(* IEC 61131-3 sources: daoli-st-library/DL_Base (part 3) *)

(* ---- FC_DL_StringRemoveWhitespace.st ---- *)
(*==============================================================================
 * 组件名称 (Component)  : FC_DL_StringRemoveWhitespace
 * 所属子库 (Sublibrary) : DL_Base
 * 当前版本 (Version)    : 1.0.0
 * 兼容性   (Platform)   : CODESYS 3.5+ / TwinCAT 3 / 汇川 InoProShop / 施耐德 Machine Expert
 *                         仅依赖 IEC 61131-3 标准字符串九函数（LEN / MID / CONCAT / FIND），零厂商私有库
 * 功能描述 (Function)   : 剔除全部空白字符（空格 0x20 / 水平制表符 0x09），压缩 HMI 报文
 *                         与条码内容（上位机常带尾随空格或制表分隔，落盘前必须净化）。
 *                         逐字符扫描，命中空白则跳过，否则追加到输出缓冲。
 *                         空白识别用字符集常量 + FIND(集合, 单字符) > 0 判定：
 *                         集合常量内含一个字面量 TAB 字符（源码直接嵌入 0x09，
 *                         不经平台转义解析，跨平台语义一致）。
 * 接口     (Interface)  : 输入 sIn 原始字符串 [-]；
 *                         输出 sOut 净化结果、uiOutLen 结果字符数 [字符]、
 *                         uiRemoved 被剔除的空白字符数 [字符]、
 *                         eErrCode 错误码（E_DL_StrWsErr）；
 *                         返回值 = bValid 净化可信标志（TRUE = sOut 可信）。
 * 边界     (Boundary)   : ① 属主边界：只剔除空格与 TAB；CR/LF 不剔除（属协议帧结构，
 *                         由 CSV 转义件负责加引号，剔除会破坏报文语义）。
 *                         ② 长度守恒校验：LEN(sIn) = uiOutLen + uiRemoved，不守恒判故障级
 *                         eInternal 并回哨兵。
 *                         ③ 全空白输入 → 输出空串、uiOutLen=0、uiRemoved=LEN(sIn)、eOk（合法）。
 *                         ④ 扫描上界取实测长度（<=255），严格有界；全索引 1 基。
 *                         ⑤ 零全局耦合（无 GVL / VAR_EXTERNAL / 物理地址）。
 * 分工声明 (Scope)      : 与 `FC_DL_StringPadLeftZeros` 分工：本件只管剔除，补位归那件；
 *                         与 `FC_DL_StringIsNumeric` 分工：净化后再做数值判定。
 * 来源标签 (Source Tag) : 原创实现（无外部代码引入）
 * 码表     (Codes)      : 本件不占用全局数字码位；出口为 BOOL + STRING + 2×UINT +
 *                         本文件内定义 enum E_DL_StrWsErr（全库唯一）。
 * 红线自检 (Redline)    : R1 ✓ 零 GVL/VAR_EXTERNAL ｜ R2 ✓ 零 %I/%Q/%M ｜ R3 ✓ 纯 IEC 61131-3
 *                         R4 ✓ 长度守恒复检 + 扫描上界钳位 + 字符集归类（无字符码强转） ｜ R5 ✓ 声明逐行同行双语注释
 *                         R6 N/A（纯函数无状态机） ｜ R7 N/A（无实例调用）
 * 修订历史 (Revision)   : 2026-11-23  v1.0.0  R77 首版（批次 B2 · 序号 6）
 * 验收向量 (Acceptance) : ① sIn=' A B '(5 字符) → sOut='AB', uiOutLen=2, uiRemoved=3, eOk, TRUE；
 *                         ② sIn='ABC' → sOut='ABC', uiOutLen=3, uiRemoved=0, eOk；
 *                         ③ sIn='   ' → sOut='', uiOutLen=0, uiRemoved=3, eOk；
 *                         ④ sIn='' → sOut='', uiOutLen=0, uiRemoved=0, eOk。
 *==============================================================================*)

(*-----------------------------------------------------------------------------
 * 枚举: E_DL_StrWsErr（空白剔除错误码，归属 DL_Base，与本件同文件，全库唯一属主）
 *----------------------------------------------------------------------------*)
TYPE E_DL_StrWsErr :
(
    eOk       := 0,   // 信息级：剔除完成 / Info: removal completed
    eInternal := 9    // 故障级：长度守恒校验失败，结果不可信 / Fault: length conservation failed, result untrustworthy
);
END_TYPE

FUNCTION FC_DL_StringRemoveWhitespace : BOOL
VAR_INPUT
    sIn : STRING(255);   // 原始字符串 [-] / Raw input string
END_VAR
VAR_OUTPUT
    sOut      : STRING(255);   // 净化结果 [-] / Sanitized result
    uiOutLen  : UINT;          // 结果字符数 [字符] / Result character count [chars]
    uiRemoved : UINT;          // 被剔除的空白字符数 [字符] / Removed whitespace character count [chars]
    eErrCode  : E_DL_StrWsErr; // 错误码出口 [-] / Error code outlet
END_VAR
VAR
    _udLen   : UDINT;        // 输入字符数（钳位后） [字符] / Input length after clamping [chars]
    _udI     : UDINT;        // 扫描位置（1 基） [-] / Scan position, 1-based
    _sCur    : STRING(255);  // 当前单字符 [-] / Current single character
    _bSkip   : BOOL;         // 当前字符是否空白 [-] / Whether current character is whitespace
    _uiDrop  : UINT;         // 剔除累加器 [字符] / Removal accumulator [chars]
END_VAR
VAR CONSTANT
    (* 空白字符集合：首个字符为空格 0x20，第二个字符为字面量 TAB 0x09（直接嵌入） *)
    (* Whitespace set: first is space 0x20, second is a literal TAB 0x09 embedded directly *)
    DL_SWS_WS_SET  : STRING(255) := '	 ';   // 空白字符集（TAB + 空格） [-] / Whitespace set, TAB plus space
    DL_SWS_LEN_MAX : UINT := 255;           // 缓冲上限（STRING(255) 契约） [字符] / Buffer ceiling [chars]
    DL_SWS_START   : UDINT := 1;            // 字符串起始位置（IEC 1 基） [-] / String start position, 1-based
    DL_SWS_ONE_LEN : UDINT := 1;            // 单字符长度常量 [字符] / Single character length constant
END_VAR

(* —— 段 0：出口预置安全值 —— *)
FC_DL_StringRemoveWhitespace := FALSE;             // 返回值预置不可信 / Return preset untrustworthy
sOut      := '';                                   // 结果哨兵空串 / Result sentinel
uiOutLen  := 0;                                    // 长度哨兵 0 / Length sentinel
uiRemoved := 0;                                    // 剔除哨兵 0 / Removal sentinel
eErrCode  := E_DL_StrWsErr.eInternal;              // 预置最严码 / Preset strictest code

(* —— 段 1：长度实测与上域钳位（缓冲可表性反算） —— *)
_udLen := LEN(sIn);                                // 输入字符数 / Input length
IF _udLen > UINT_TO_UDINT(DL_SWS_LEN_MAX) THEN
    _udLen := UINT_TO_UDINT(DL_SWS_LEN_MAX);       // 超上限钳位 / Clamp to ceiling
END_IF

(* —— 段 2：空串早退（合法零结果） —— *)
IF _udLen = 0 THEN
    eErrCode := E_DL_StrWsErr.eOk;                 // 信息级成功 / Info success
    FC_DL_StringRemoveWhitespace := TRUE;
    RETURN;
END_IF

(* —— 段 3：逐字符扫描与选择性追加 —— *)
_uiDrop := 0;                                      // 剔除累加器清零 / Clear removal accumulator
_udI    := DL_SWS_START;                           // 起算位置 1 / Start at position one
sOut    := '';                                     // 输出缓冲显式清空 / Explicitly clear output buffer
WHILE _udI <= _udLen DO
    _sCur  := MID(sIn, DL_SWS_ONE_LEN, _udI);      // 取第 i 个字符（1 基） / Take i-th character, 1-based
    _bSkip := (FIND(DL_SWS_WS_SET, _sCur) > 0);    // 命中空白集合即跳过 / Skip when hit whitespace set
    IF _bSkip THEN
        _uiDrop := _uiDrop + 1;                    // 剔除累加 / Accumulate removal
    ELSE
        sOut := CONCAT(sOut, _sCur);               // 非空白追加 / Append non-whitespace character
    END_IF
    _udI := _udI + 1;                              // 位置步进 / Advance position
END_WHILE

(* —— 段 4：长度守恒复检（输入长度 = 保留 + 剔除） —— *)
uiOutLen  := UDINT_TO_UINT(LEN(sOut));             // 结果字符数 / Result length
uiRemoved := _uiDrop;                              // 剔除字符数 / Removed count
IF (UDINT_TO_UINT(_udLen) <> (uiOutLen + uiRemoved)) THEN
    sOut      := '';                               // 守恒失败回哨兵 / Conservation failed: sentinel
    uiOutLen  := 0;
    uiRemoved := 0;
    eErrCode  := E_DL_StrWsErr.eInternal;          // 故障级码 / Fault-level code
    RETURN;                                        // 返回 FALSE 保持 / Keep return FALSE
END_IF

(* —— 段 5：成功出口 —— *)
eErrCode := E_DL_StrWsErr.eOk;                     // 信息级成功 / Info success
FC_DL_StringRemoveWhitespace := TRUE;              // 净化可信 / Sanitization trustworthy

END_FUNCTION

(* ---- FC_DL_StringRepeat.st ---- *)
(*==============================================================================
 * 组件名称 (Component)  : FC_DL_StringRepeat
 * 所属子库 (Sublibrary) : DL_Base
 * 当前版本 (Version)    : 1.0.0
 * 兼容性   (Platform)   : CODESYS 3.5+ / TwinCAT 3 / 汇川 InoProShop / 施耐德 Machine Expert
 *                         仅依赖 IEC 61131-3 标准字符串九函数（LEN / CONCAT），零厂商私有库
 * 功能描述 (Function)   : 按次数重复拼接（分隔线 "-----"、占位符 "<><><>"、缩进填充）。
 *                         先算缓冲可容最大重复次数 = 255 DIV LEN(sIn)（分母已判零，
 *                         结构性无除零），再与请求次数比较：请求超限则按最大可容次数
 *                         截断并置 bTruncated / eTruncated（信息级，结果仍可信）；
 *                         请求次数为 0 或输入空串时输出空串。
 * 接口     (Interface)  : 输入 sIn 基元字符串 [-]、uiCount 请求重复次数 [次]；
 *                         输出 sOut 拼接结果、uiOutLen 结果字符数 [字符]、
 *                         uiApplied 实际生效次数 [次]、bTruncated 截断回执、
 *                         eErrCode 错误码（E_DL_StrRepErr）；
 *                         返回值 = bValid 拼接可信标志（TRUE = sOut 可信）。
 * 边界     (Boundary)   : ① 属主边界：只做整串重复拼接，不做单字符补位（补位归
 *                         FC_DL_StringPadLeftZeros）、不做截断加标记（归 TruncEllipsis）。
 *                         ② 除零防御：先判 LEN(sIn)=0 并早退，后才做 255 DIV LEN(sIn)。
 *                         ③ 缓冲保护：结果长度恒 <= 255（生效次数 = 255 DIV 基元长度）。
 *                         ④ uiCount=0 → 输出空串、uiApplied=0、eOk（合法零次）。
 *                         ⑤ 零全局耦合（无 GVL / VAR_EXTERNAL / 物理地址）。
 * 分工声明 (Scope)      : 与 `FC_DL_StringPadLeftZeros` 分工：定长补位归那件、
 *                         次数重复归本件；与 `FC_DL_StringTruncEllipsis` 无调用关系。
 * 来源标签 (Source Tag) : 原创实现（无外部代码引入）
 * 码表     (Codes)      : 本件不占用全局数字码位；出口为 BOOL + STRING + 3×UINT +
 *                         本文件内定义 enum E_DL_StrRepErr（全库唯一）。
 * 红线自检 (Redline)    : R1 ✓ 零 GVL/VAR_EXTERNAL ｜ R2 ✓ 零 %I/%Q/%M ｜ R3 ✓ 纯 IEC 61131-3
 *                         R4 ✓ 除零前置判零 + 缓冲上限反算 + 循环次数有界 ｜ R5 ✓ 声明逐行同行双语注释
 *                         R6 N/A（纯函数无状态机） ｜ R7 N/A（无实例调用）
 * 修订历史 (Revision)   : 2026-11-23  v1.0.0  R77 首版（批次 B2 · 序号 8）
 * 验收向量 (Acceptance) : ① sIn='AB', uiCount=3 → sOut='ABABAB', uiOutLen=6, uiApplied=3,
 *                         bTruncated=FALSE, eOk, TRUE；
 *                         ② sIn='AB', uiCount=0 → sOut='', uiOutLen=0, uiApplied=0, eOk, TRUE；
 *                         ③ sIn='', uiCount=5 → sOut='', uiOutLen=0, uiApplied=0, eOk, TRUE；
 *                         ④ sIn='X'（1 字符）, uiCount=300 → 生效 255 次，sOut 长度 255,
 *                         bTruncated=TRUE, eTruncated；
 *                         ⑤ sIn='AB', uiCount=200 → 255 DIV 2 = 127 → uiApplied=127,
 *                         长度 254, bTruncated=TRUE。
 *==============================================================================*)

(*-----------------------------------------------------------------------------
 * 枚举: E_DL_StrRepErr（重复拼接错误码，归属 DL_Base，与本件同文件，全库唯一属主）
 *----------------------------------------------------------------------------*)
TYPE E_DL_StrRepErr :
(
    eOk        := 0,   // 信息级：按请求次数完成 / Info: completed as requested
    eTruncated := 1    // 信息级：超缓冲上限已按最大可容次数截断 / Info: truncated to max fitting repeat count
);
END_TYPE

FUNCTION FC_DL_StringRepeat : BOOL
VAR_INPUT
    sIn     : STRING(255);   // 基元字符串 [-] / Unit string to repeat
    uiCount : UINT;          // 请求重复次数 [次] / Requested repeat count [times]
END_VAR
VAR_OUTPUT
    sOut       : STRING(255); // 拼接结果 [-] / Concatenated result
    uiOutLen   : UINT;        // 结果字符数 [字符] / Result character count [chars]
    uiApplied  : UINT;        // 实际生效次数 [次] / Applied repeat count [times]
    bTruncated : BOOL;        // 截断回执（信息级） [-] / Truncation receipt, info level
    eErrCode   : E_DL_StrRepErr; // 错误码出口 [-] / Error code outlet
END_VAR
VAR
    _udUnitLen : UDINT;       // 基元字符数 [字符] / Unit string length [chars]
    _udMaxRep  : UDINT;       // 缓冲可容最大重复次数 [次] / Max fitting repeat count [times]
    _uiEff     : UINT;        // 生效重复次数 [次] / Effective repeat count [times]
    _uiLoop    : UINT;        // 循环计数器 [-] / Loop counter
END_VAR
VAR CONSTANT
    DL_SRE_LEN_MAX : UINT := 255;    // 缓冲上限（STRING(255) 契约） [字符] / Buffer ceiling [chars]
    DL_SRE_ONE_LEN : UDINT := 1;     // 单字符长度常量 [字符] / Single character length constant
END_VAR

(* —— 段 0：出口预置安全值 —— *)
FC_DL_StringRepeat := FALSE;                       // 返回值预置无效 / Return preset invalid
sOut       := '';                                  // 结果哨兵空串 / Result sentinel
uiOutLen   := 0;                                   // 长度哨兵 0 / Length sentinel
uiApplied  := 0;                                   // 生效次数哨兵 0 / Applied count sentinel
bTruncated := FALSE;                               // 截断回执预置无 / Truncation receipt preset false
eErrCode   := E_DL_StrRepErr.eTruncated;           // 预置最严码（本件仅信息级码） / Preset strictest code

(* —— 段 1：基元长度实测（除零防御前置：先判零后做除法） —— *)
_udUnitLen := LEN(sIn);                            // 基元字符数 / Unit length
IF _udUnitLen = 0 THEN
    eErrCode := E_DL_StrRepErr.eOk;                // 空基元合法（零结果） / Empty unit is legal, zero result
    FC_DL_StringRepeat := TRUE;                    // 结果可信 / Result trustworthy
    RETURN;                                        // 早退，彻底规避 255 DIV 0 / Early exit, avoids division by zero entirely
END_IF

(* —— 段 2：请求次数为零早退（合法零结果） —— *)
IF uiCount = 0 THEN
    eErrCode := E_DL_StrRepErr.eOk;                // 零次合法 / Zero repeats legal
    FC_DL_StringRepeat := TRUE;
    RETURN;
END_IF

(* —— 段 3：缓冲可容最大重复次数反算（分母已确非零） —— *)
_udMaxRep := UINT_TO_UDINT(DL_SRE_LEN_MAX) / _udUnitLen;  // 255 DIV 基元长度 / Integer division by unit length
IF _udMaxRep < DL_SRE_ONE_LEN THEN
    _udMaxRep := DL_SRE_ONE_LEN;                   // 基元本身已占满缓冲：至少一次 / Unit already fills buffer: at least once
END_IF

(* —— 段 4：请求次数与可容次数比较（超限则截断并回执） —— *)
IF UINT_TO_UDINT(uiCount) > _udMaxRep THEN
    _uiEff     := UDINT_TO_UINT(_udMaxRep);         // 收敛到最大可容次数 / Converge to max fitting count
    bTruncated := TRUE;                            // 截断回执 / Truncation receipt
    eErrCode   := E_DL_StrRepErr.eTruncated;       // 信息级截断码 / Info truncation code
ELSE
    _uiEff     := uiCount;                         // 按请求次数生效 / Apply requested count
    bTruncated := FALSE;
    eErrCode   := E_DL_StrRepErr.eOk;              // 信息级成功 / Info success
END_IF

(* —— 段 5：循环拼接（次数已收敛，循环严格有界） —— *)
sOut := '';                                        // 输出缓冲显式清空 / Explicitly clear output buffer
IF _uiEff > 0 THEN
    FOR _uiLoop := 1 TO _uiEff DO
        sOut := CONCAT(sOut, sIn);                 // 每次追加一个基元 / Append one unit per iteration
    END_FOR;
END_IF

(* —— 段 6：结果复检（长度 = 基元长度 × 生效次数，且不得超缓冲） —— *)
uiOutLen  := UDINT_TO_UINT(LEN(sOut));             // 实测结果长度 / Measured result length
uiApplied := _uiEff;                               // 导出生效次数 / Export applied count
IF uiOutLen > DL_SRE_LEN_MAX THEN
    sOut      := '';                               // 超缓冲回哨兵 / Over buffer: sentinel
    uiOutLen  := 0;
    uiApplied := 0;
    eErrCode  := E_DL_StrRepErr.eTruncated;        // 保持信息级码（本件无故障级码位） / Keep info-level code
    RETURN;
END_IF

FC_DL_StringRepeat := TRUE;                        // 拼接有效 / Concatenation valid

END_FUNCTION

(* ---- FC_DL_StringReverse.st ---- *)
(*==============================================================================
 * 组件名称 (Component)  : FC_DL_StringReverse
 * 所属子库 (Sublibrary) : DL_Base
 * 当前版本 (Version)    : 1.0.0
 * 兼容性   (Platform)   : CODESYS 3.5+ / TwinCAT 3 / 汇川 InoProShop / 施耐德 Machine Expert
 *                         仅依赖 IEC 61131-3 标准字符串九函数（LEN / MID / CONCAT），零厂商私有库
 * 功能描述 (Function)   : 字符串反转（回文校验 / 字节序调试 / 低位在前的编码还原）。
 *                         自尾向头逐字符取 MID(sIn,1,i) 并 CONCAT 拼接；用 WHILE
 *                         递减计数，UDINT 计数到 0 自然终止，结构上无下溢路径。
 *                         输出长度恒等于输入长度（不做任何增删）。
 * 接口     (Interface)  : 输入 sIn 原始字符串 [-]；
 *                         输出 sOut 反转结果、uiOutLen 结果字符数 [字符]、
 *                         eErrCode 错误码（E_DL_StrRevErr）；
 *                         返回值 = bValid 反转可信标志（TRUE = sOut 可信）。
 * 边界     (Boundary)   : ① 属主边界：只做整串反转，不做大小写折叠、不做子串反转。
 *                         ② 长度 > 255 时按缓冲上限 255 截断尾部（保证输出可表），
 *                         回执 eClampLen（信息级），bTruncated 置位。
 *                         ③ 空串合法，输出空串、uiOutLen=0、eOk。
 *                         ④ 计数递减用 `IF _udI > 0` 前置判定，杜绝 UDINT 0-1 下溢。
 *                         ⑤ 零全局耦合（无 GVL / VAR_EXTERNAL / 物理地址）。
 * 分工声明 (Scope)      : 与 `FC_DL_StringCompareNatural` 分工：反转只做位序重排，
 *                         不做序比较；回文判定由调用方对 sIn 与 sOut 比较完成。
 * 来源标签 (Source Tag) : 原创实现（无外部代码引入）
 * 码表     (Codes)      : 本件不占用全局数字码位；出口为 BOOL + STRING + UINT +
 *                         本文件内定义 enum E_DL_StrRevErr（全库唯一）。
 * 红线自检 (Redline)    : R1 ✓ 零 GVL/VAR_EXTERNAL ｜ R2 ✓ 零 %I/%Q/%M ｜ R3 ✓ 纯 IEC 61131-3
 *                         R4 ✓ 递减计数下溢防护 + 长度钳位 ｜ R5 ✓ 声明逐行同行双语注释
 *                         R6 N/A（纯函数无状态机） ｜ R7 N/A（无实例调用）
 * 修订历史 (Revision)   : 2026-11-23  v1.0.0  R77 首版（批次 B2 · 序号 4）
 * 验收向量 (Acceptance) : ① sIn='ABC' → sOut='CBA', uiOutLen=3, eOk, TRUE；
 *                         ② sIn='ABBA' → sOut='ABBA'（回文自反）, uiOutLen=4；
 *                         ③ sIn='' → sOut='', uiOutLen=0, eOk, TRUE；
 *                         ④ sIn='12345' → sOut='54321'。
 *==============================================================================*)

(*-----------------------------------------------------------------------------
 * 枚举: E_DL_StrRevErr（字符串反转错误码，归属 DL_Base，与本件同文件，全库唯一属主）
 *----------------------------------------------------------------------------*)
TYPE E_DL_StrRevErr :
(
    eOk       := 0,   // 信息级：反转完成 / Info: reversal completed
    eClampLen := 1    // 信息级：长度超缓冲上限已截断 / Info: length clamped to buffer ceiling
);
END_TYPE

FUNCTION FC_DL_StringReverse : BOOL
VAR_INPUT
    sIn : STRING(255);   // 原始字符串 [-] / Raw input string
END_VAR
VAR_OUTPUT
    sOut      : STRING(255);   // 反转结果 [-] / Reversed result
    uiOutLen  : UINT;          // 结果字符数 [字符] / Result character count [chars]
    bTruncated: BOOL;          // 截断回执（信息级） [-] / Truncation receipt, info level
    eErrCode  : E_DL_StrRevErr; // 错误码出口 [-] / Error code outlet
END_VAR
VAR
    _udLen : UDINT;       // 生效字符数（钳位后） [字符] / Effective character count after clamping [chars]
    _udI   : UDINT;       // 逆序扫描位置（1 基） [-] / Reverse scan position, 1-based
END_VAR
VAR CONSTANT
    DL_SRV_LEN_MAX : UINT := 255;    // 缓冲上限（STRING(255) 契约） [字符] / Buffer ceiling [chars]
    DL_SRV_ONE_LEN : UDINT := 1;     // 单字符长度常量 [字符] / Single character length constant [chars]
END_VAR

(* —— 段 0：出口预置安全值 —— *)
FC_DL_StringReverse := FALSE;                      // 返回值预置无效 / Return preset invalid
sOut       := '';                                  // 结果哨兵空串 / Result sentinel
uiOutLen   := 0;                                   // 长度哨兵 0 / Length sentinel
bTruncated := FALSE;                               // 截断回执预置无 / Truncation receipt preset false
eErrCode   := E_DL_StrRevErr.eClampLen;            // 预置最严码（本件仅信息级码） / Preset strictest code

(* —— 段 1：长度实测与上域钳位（缓冲可表性反算） —— *)
_udLen := LEN(sIn);                                // 输入字符数 / Input length
IF _udLen > UINT_TO_UDINT(DL_SRV_LEN_MAX) THEN
    _udLen     := UINT_TO_UDINT(DL_SRV_LEN_MAX);   // 超上限截断尾部 / Truncate tail beyond ceiling
    bTruncated := TRUE;                            // 截断回执 / Truncation receipt
    eErrCode   := E_DL_StrRevErr.eClampLen;        // 信息级钳位码 / Info clamp code
ELSE
    eErrCode   := E_DL_StrRevErr.eOk;              // 信息级成功 / Info success
END_IF

(* —— 段 2：空串早退（合法零结果） —— *)
IF _udLen = 0 THEN
    FC_DL_StringReverse := TRUE;                   // 空串反转合法 / Empty reversal legal
    RETURN;
END_IF

(* —— 段 3：逆序拼接（前置 >0 判定，杜绝 UDINT 下溢） —— *)
sOut := MID(sIn, DL_SRV_ONE_LEN, _udLen);          // 以末字符起头 / Start with last character
_udI := _udLen - 1;                                // 自倒数第二位起（>=1 由段 2 保证 len>=1） / Start from second last
WHILE _udI > 0 DO
    sOut := CONCAT(sOut, MID(sIn, DL_SRV_ONE_LEN, _udI));  // 逐个前置字符追加 / Append next character from tail
    _udI := _udI - 1;                              // 位置递减，条件 >0 保证不下溢 / Decrement, guarded by >0
END_WHILE

(* —— 段 4：结果复检（长度守恒） —— *)
uiOutLen := UDINT_TO_UINT(LEN(sOut));              // 实测结果长度 / Measured result length
IF uiOutLen <> UDINT_TO_UINT(_udLen) THEN
    sOut     := '';                                // 长度不守恒回哨兵 / Length not conserved: sentinel
    uiOutLen := 0;
    eErrCode := E_DL_StrRevErr.eClampLen;          // 保持信息级码（本件无故障级码位） / Keep info-level code
END_IF

FC_DL_StringReverse := TRUE;                       // 反转有效（含截断情形） / Reversal valid, truncation included

END_FUNCTION

(* ---- FC_DL_StringSplitPair.st ---- *)
(*==============================================================================
 * 组件名称 (Component)  : FC_DL_StringSplitPair
 * 所属子库 (Sublibrary) : DL_Base
 * 当前版本 (Version)    : 1.0.0
 * 兼容性   (Platform)   : CODESYS 3.5+ / TwinCAT 3 / 汇川 InoProShop / 施耐德 Machine Expert
 *                         仅依赖 IEC 61131-3 标准字符串九函数（LEN / MID / FIND），零厂商私有库
 * 功能描述 (Function)   : key=value 单对拆分（HMI 参数设置报文 "Speed=1500" 解析）。
 *                         以首个分隔符位置为界：左侧为键、右侧为值（值可含分隔符，
 *                         故只按首个分隔符切分）。缺分隔符、空键均置无效回执（返回 FALSE），
 *                         空值合法（代表「置空」语义，回执 bHasValue=FALSE 但不判故障）。
 *                         分隔符为可配字符串（默认 '='），支持 ':=' / '->' 等双字符分隔。
 * 接口     (Interface)  : 输入 sIn 待拆分字符串 [-]、sSep 分隔符（空串回落 '='）[-]；
 *                         输出 sKey 键、sValue 值、uiKeyLen 键长 [字符]、uiValueLen 值长 [字符]、
 *                         bHasValue 是否存在值段、eErrCode 错误码（E_DL_StrSplitErr）；
 *                         返回值 = bValid 拆分有效标志（TRUE = sKey/sValue 可信）。
 * 边界     (Boundary)   : ① 属主边界：只拆单对，不遍历多对、不去引号、不做类型转换。
 *                         ② 缺分隔符 → 故障级 eNoSeparator，sKey=sIn 原样、sValue=''、返回 FALSE。
 *                         ③ 分隔符在首位（空键）→ 故障级 eEmptyKey，sKey=''、sValue=右段。
 *                         ④ 分隔符在末位（空值）→ 信息级 eEmptyValue，bHasValue=FALSE、返回 TRUE。
 *                         ⑤ MID 起算位置 = 分隔符位置 + 1，且仅当剩余长度 >= 1 时才取，
 *                         结构上无 0 长度 / 0 位置取值路径。
 *                         ⑥ 零全局耦合（无 GVL / VAR_EXTERNAL / 物理地址）。
 * 分工声明 (Scope)      : 与 `FC_DL_StringCountChar` 分工：计数归那件、拆分归本件；
 *                         与 `FC_DL_StringCsvFieldEscape` 分工：CSV 转义归那件。
 * 来源标签 (Source Tag) : 原创实现（无外部代码引入）
 * 码表     (Codes)      : 本件不占用全局数字码位；出口为 BOOL + 2×STRING + 2×UINT +
 *                         本文件内定义 enum E_DL_StrSplitErr（全库唯一）。
 * 红线自检 (Redline)    : R1 ✓ 零 GVL/VAR_EXTERNAL ｜ R2 ✓ 零 %I/%Q/%M ｜ R3 ✓ 纯 IEC 61131-3
 *                         R4 ✓ 分隔符缺失/空键域闸 + 取值位置下限保护 ｜ R5 ✓ 声明逐行同行双语注释
 *                         R6 N/A（纯函数无状态机） ｜ R7 N/A（无实例调用）
 * 修订历史 (Revision)   : 2026-11-23  v1.0.0  R77 首版（批次 B2 · 序号 7）
 * 验收向量 (Acceptance) : ① sIn='Speed=1500', sSep='=' → sKey='Speed', sValue='1500',
 *                         uiKeyLen=5, uiValueLen=4, bHasValue=TRUE, eOk, TRUE；
 *                         ② sIn='Speed1450', sSep='=' → bFound 无效：返回 FALSE, eNoSeparator, sValue=''；
 *                         ③ sIn='=1500' → 返回 FALSE, eEmptyKey, sKey='';
 *                         ④ sIn='Speed=' → sKey='Speed', sValue='', bHasValue=FALSE,
 *                         返回 TRUE, eEmptyValue；
 *                         ⑤ sIn='A=B=C' → sKey='A', sValue='B=C'（只按首个分隔符切分）；
 *                         ⑥ sIn='', sSep='=' → 返回 FALSE, eNoSeparator。
 *==============================================================================*)

(*-----------------------------------------------------------------------------
 * 枚举: E_DL_StrSplitErr（key=value 拆分错误码，归属 DL_Base，与本件同文件，全库唯一属主）
 * 分级: eEmptyValue 为信息级（返回 TRUE）；eNoSeparator / eEmptyKey 为故障级（返回 FALSE）。
 *----------------------------------------------------------------------------*)
TYPE E_DL_StrSplitErr :
(
    eOk          := 0,   // 信息级：键值均非空，拆分完成 / Info: both key and value non-empty
    eEmptyValue  := 1,   // 信息级：值段为空（置空语义） / Info: empty value section
    eNoSeparator := 2,   // 故障级：未找到分隔符 / Fault: separator not found
    eEmptyKey    := 3    // 故障级：分隔符在首位，键为空 / Fault: separator at head, empty key
);
END_TYPE

FUNCTION FC_DL_StringSplitPair : BOOL
VAR_INPUT
    sIn  : STRING(255);   // 待拆分字符串 [-] / String to split
    sSep : STRING(255);   // 分隔符（空串回落 '='） [-] / Separator, empty falls back to '='
END_VAR
VAR_OUTPUT
    sKey       : STRING(255); // 键段 [-] / Key section
    sValue     : STRING(255); // 值段 [-] / Value section
    uiKeyLen   : UINT;        // 键字符数 [字符] / Key character count [chars]
    uiValueLen : UINT;        // 值字符数 [字符] / Value character count [chars]
    bHasValue  : BOOL;        // 是否存在值段 [-] / Whether value section exists
    eErrCode   : E_DL_StrSplitErr; // 错误码出口 [-] / Error code outlet
END_VAR
VAR
    _sSepUse  : STRING(255);  // 生效分隔符 [-] / Effective separator
    _udLen    : UDINT;        // 输入字符数（钳位后） [字符] / Input length after clamping [chars]
    _udPos    : UDINT;        // 分隔符位置（1 基，0 = 未找到） [-] / Separator position, 0 means not found
    _udRemain : UDINT;        // 分隔符右侧剩余字符数 [字符] / Remaining characters after separator [chars]
    _udStart  : UDINT;        // 值段起算位置（1 基） [-] / Value section start position, 1-based
END_VAR
VAR CONSTANT
    DL_SSP_SEP_DFLT : STRING(255) := '=';   // 默认分隔符 [-] / Default separator
    DL_SSP_LEN_MAX  : UINT := 255;          // 缓冲上限（STRING(255) 契约） [字符] / Buffer ceiling [chars]
    DL_SSP_START    : UDINT := 1;           // 字符串起始位置（IEC 1 基） [-] / String start position, 1-based
END_VAR

(* —— 段 0：出口预置安全值 —— *)
FC_DL_StringSplitPair := FALSE;                    // 返回值预置无效 / Return preset invalid
sKey       := '';                                  // 键哨兵空串 / Key sentinel
sValue     := '';                                  // 值哨兵空串 / Value sentinel
uiKeyLen   := 0;                                   // 键长哨兵 0 / Key length sentinel
uiValueLen := 0;                                   // 值长哨兵 0 / Value length sentinel
bHasValue  := FALSE;                               // 值段存在性预置无 / Value presence preset false
eErrCode   := E_DL_StrSplitErr.eNoSeparator;       // 预置最严码 / Preset strictest code

(* —— 段 1：分隔符归一（空串回落默认 '='） —— *)
IF LEN(sSep) = 0 THEN
    _sSepUse := DL_SSP_SEP_DFLT;                   // 回落默认分隔符 / Fall back to default separator
ELSE
    _sSepUse := sSep;                              // 使用调用方给定分隔符 / Use caller-supplied separator
END_IF

(* —— 段 2：输入长度实测与上域钳位 —— *)
_udLen := LEN(sIn);                                // 输入字符数 / Input length
IF _udLen > UINT_TO_UDINT(DL_SSP_LEN_MAX) THEN
    _udLen := UINT_TO_UDINT(DL_SSP_LEN_MAX);       // 超上限钳位 / Clamp to ceiling
END_IF

(* —— 段 3：定位首个分隔符（FIND 返回 0 表示未找到） —— *)
_udPos := FIND(sIn, _sSepUse);                     // 首个分隔符位置（1 基） / First separator position, 1-based

(* —— 段 4：缺分隔符早退（故障级：整体原样回键，值置空） —— *)
IF _udPos = 0 THEN
    sKey     := sIn;                               // 原样回键便于调用方诊断 / Echo input to key for diagnosis
    uiKeyLen := UDINT_TO_UINT(LEN(sKey));          // 键长实测 / Measured key length
    sValue   := '';                                // 值置空 / Value cleared
    eErrCode := E_DL_StrSplitErr.eNoSeparator;     // 故障级码 / Fault-level code
    RETURN;                                        // 返回 FALSE 保持 / Keep return FALSE
END_IF

(* —— 段 5：空键闸（分隔符在首位） —— *)
IF _udPos = DL_SSP_START THEN
    sKey     := '';                                // 键为空 / Empty key
    _udRemain := _udLen - _udPos;                  // 右侧剩余长度 / Remaining length on the right
    IF _udRemain >= DL_SSP_START THEN
        sValue     := MID(sIn, _udRemain, _udPos + DL_SSP_START);  // 取分隔符之后全部字符 / Take all after separator
        uiValueLen := UDINT_TO_UINT(_udRemain);
        bHasValue  := TRUE;
    END_IF
    eErrCode := E_DL_StrSplitErr.eEmptyKey;        // 故障级码 / Fault-level code
    RETURN;                                        // 返回 FALSE 保持 / Keep return FALSE
END_IF

(* —— 段 6：键段提取（位置 1 起，长度 = 分隔符位置 - 1 >= 1） —— *)
sKey     := MID(sIn, _udPos - DL_SSP_START, DL_SSP_START);   // 分隔符左侧 / Left of separator
uiKeyLen := UDINT_TO_UINT(LEN(sKey));              // 键长实测 / Measured key length

(* —— 段 7：值段提取（起算位置 = 分隔符位置 + 1，仅剩余 >= 1 时取） —— *)
_udRemain := _udLen - _udPos;                      // 右侧剩余长度 / Remaining length on the right
IF _udRemain >= DL_SSP_START THEN
    _udStart   := _udPos + DL_SSP_START;           // 值段起算位置 / Value start position
    sValue     := MID(sIn, _udRemain, _udStart);   // 取右侧全部字符 / Take all characters on the right
    uiValueLen := UDINT_TO_UINT(LEN(sValue));      // 值长实测 / Measured value length
    bHasValue  := TRUE;                            // 存在值段 / Value section exists
    eErrCode   := E_DL_StrSplitErr.eOk;            // 信息级成功 / Info success
ELSE
    sValue     := '';                              // 分隔符在末位：值段为空 / Separator at tail: empty value
    uiValueLen := 0;
    bHasValue  := FALSE;
    eErrCode   := E_DL_StrSplitErr.eEmptyValue;    // 信息级：置空语义 / Info: clear semantics
END_IF

(* —— 段 8：键长复检（键不得为空，否则判内部不一致） —— *)
IF uiKeyLen = 0 THEN
    sKey     := '';                                // 回哨兵 / Back to sentinel
    sValue   := '';
    eErrCode := E_DL_StrSplitErr.eEmptyKey;        // 故障级码 / Fault-level code
    RETURN;
END_IF

FC_DL_StringSplitPair := TRUE;                     // 拆分有效 / Split valid

END_FUNCTION

(* ---- FC_DL_StringTruncEllipsis.st ---- *)
(*==============================================================================
 * 组件名称 (Component)  : FC_DL_StringTruncEllipsis
 * 所属子库 (Sublibrary) : DL_Base
 * 当前版本 (Version)    : 1.0.0
 * 兼容性   (Platform)   : CODESYS 3.5+ / TwinCAT 3 / 汇川 InoProShop / 施耐德 Machine Expert
 *                         仅依赖 IEC 61131-3 标准字符串九函数（LEN / MID / CONCAT），零厂商私有库
 * 功能描述 (Function)   : 超长截断并补省略标记（HMI 单行显示 / 报警摘要压缩）。
 *                         sIn 长度不超过 uiMaxLen 时原样返回；超长时保留前
 *                         (uiMaxLen - LEN(sMark)) 个字符并追加省略标记，最终长度
 *                         恒等于 uiMaxLen（标记有余量时）；标记本身已占满目标长度时
 *                         退化为纯截断（无标记空间）并回执 eTruncNoMark。
 *                         返回实际写入字符数 uiOutLen，供调用方做定宽对齐。
 * 接口     (Interface)  : 输入 sIn 原始字符串 [-]、uiMaxLen 目标最大长度（含标记）[字符]、
 *                         sMark 省略标记（空串则纯截断）[-]；
 *                         输出 sOut 结果字符串、uiOutLen 实际字符数 [字符]、
 *                         bTruncated 截断回执、eErrCode 错误码（E_DL_StrTruncErr）；
 *                         返回值 = bValid 输出可信标志（TRUE = sOut 可信）。
 * 边界     (Boundary)   : ① 属主边界：只做截断 + 单标记追加，不做补位、不剔除空白。
 *                         ② uiMaxLen 合法域 1..255；> 255 钳位至 255 并置 eClampLen；
 *                         < 1 判故障级 eInvalidParam（无法产出有效结果）。
 *                         ③ 标记长度 >= uiMaxLen 时无标记余量，退化为 MID(sIn,uiMaxLen,1)
 *                         纯截断，回执 eTruncNoMark（信息级）。
 *                         ④ 全索引 1 基，截断起算位置恒 >= 1（keep >= 1 由分支保证）。
 *                         ⑤ 零全局耦合（无 GVL / VAR_EXTERNAL / 物理地址）。
 * 分工声明 (Scope)      : 与 `FC_DL_StringPadLeftZeros` 分工：补位归那件、截断归本件，
 *                         两件互不调用；与 `FC_DL_StringRepeat` 无交集。
 * 来源标签 (Source Tag) : 原创实现（无外部代码引入）
 * 码表     (Codes)      : 本件不占用全局数字码位；出口为 BOOL + STRING + UINT +
 *                         本文件内定义 enum E_DL_StrTruncErr（全库唯一）。
 * 红线自检 (Redline)    : R1 ✓ 零 GVL/VAR_EXTERNAL ｜ R2 ✓ 零 %I/%Q/%M ｜ R3 ✓ 纯 IEC 61131-3
 *                         R4 ✓ 长度域闸 + 双侧钳位 + 起算位置下限保证 ｜ R5 ✓ 声明逐行同行双语注释
 *                         R6 N/A（纯函数无状态机） ｜ R7 N/A（无实例调用）
 * 修订历史 (Revision)   : 2026-11-23  v1.0.0  R77 首版（批次 B2 · 序号 2）
 * 验收向量 (Acceptance) : ① sIn='ABCDEFGH'（8 字符）, uiMaxLen=6, sMark='...' →
 *                         keep=3 → sOut='ABC...'（6 字符）, uiOutLen=6, bTruncated=TRUE, eOk；
 *                         ② sIn='ABC', uiMaxLen=6 → sOut='ABC'（原样）, uiOutLen=3,
 *                         bTruncated=FALSE, eOk；
 *                         ③ sIn='ABCDEFGH', uiMaxLen=3, sMark='...' → 标记占满 →
 *                         sOut='ABC', uiOutLen=3, bTruncated=TRUE, eTruncNoMark；
 *                         ④ uiMaxLen=0 → 返回 FALSE, sOut='', eInvalidParam。
 *==============================================================================*)

(*-----------------------------------------------------------------------------
 * 枚举: E_DL_StrTruncErr（截断错误码，归属 DL_Base，与本件同文件，全库唯一属主）
 *----------------------------------------------------------------------------*)
TYPE E_DL_StrTruncErr :
(
    eOk           := 0,   // 信息级：标记有余量，已按目标长度截断 / Info: truncated to target length with mark
    eTruncNoMark  := 1,   // 信息级：标记无余量，退化为纯截断 / Info: no room for mark, plain truncation
    eClampLen     := 2,   // 信息级：目标长度超缓冲上限已钳位 / Info: target length clamped to buffer ceiling
    eInvalidParam := 3    // 故障级：目标长度小于 1，无法产出有效结果 / Fault: target length below 1
);
END_TYPE

FUNCTION FC_DL_StringTruncEllipsis : BOOL
VAR_INPUT
    sIn      : STRING(255);   // 原始字符串 [-] / Raw input string
    uiMaxLen : UINT;          // 目标最大长度（含省略标记），合法域 1..255 [字符] / Target max length including mark, domain 1..255 [chars]
    sMark    : STRING(255);   // 省略标记（空串则退化为纯截断） [-] / Ellipsis mark, empty means plain truncation
END_VAR
VAR_OUTPUT
    sOut       : STRING(255); // 截断结果字符串 [-] / Truncated result string
    uiOutLen   : UINT;        // 实际写入字符数 [字符] / Actual written character count [chars]
    bTruncated : BOOL;        // 截断回执（信息级） [-] / Truncation receipt, info level
    eErrCode   : E_DL_StrTruncErr; // 错误码出口 [-] / Error code outlet
END_VAR
VAR
    _udInLen  : UDINT;        // 输入字符数（LEN 原生宽度） [字符] / Input length in native LEN width [chars]
    _udMarkLen: UDINT;        // 标记字符数 [字符] / Mark length [chars]
    _udKeep   : UDINT;        // 需保留的正文前缀字符数 [字符] / Number of leading text characters kept [chars]
    _udCopy   : UDINT;        // 实际拷贝字符数（钳位后） [字符] / Actual copied characters after clamping [chars]
END_VAR
VAR CONSTANT
    DL_STE_LEN_MAX  : UINT := 255;   // 缓冲上限（STRING(255) 契约） [字符] / Buffer ceiling per STRING(255) [chars]
    DL_STE_LEN_MIN  : UINT := 1;     // 目标长度下限 [字符] / Target length lower bound [chars]
    DL_STE_START    : UDINT := 1;    // 字符串起始位置（IEC 1 基） [-] / String start position, IEC 1-based
END_VAR

(* —— 段 0：出口预置安全值 —— *)
FC_DL_StringTruncEllipsis := FALSE;               // 返回值预置无效 / Return preset invalid
sOut       := '';                                  // 结果哨兵空串 / Result sentinel
uiOutLen   := 0;                                   // 长度哨兵 0 / Length sentinel
bTruncated := FALSE;                               // 截断回执预置无 / Truncation receipt preset false
eErrCode   := E_DL_StrTruncErr.eInvalidParam;      // 预置最严码 / Preset strictest code

(* —— 段 1：目标长度下域闸 —— *)
IF uiMaxLen < DL_STE_LEN_MIN THEN
    RETURN;                                        // 目标长度非法：保持故障码与哨兵 / Illegal target length
END_IF

(* —— 段 2：目标长度上域钳位（缓冲可表性反算） —— *)
IF uiMaxLen > DL_STE_LEN_MAX THEN
    uiMaxLen := DL_STE_LEN_MAX;                    // 钳位至缓冲上限 / Clamp to buffer ceiling
    eErrCode := E_DL_StrTruncErr.eClampLen;        // 信息级钳位码 / Info clamp code
END_IF

(* —— 段 3：实测长度（标准函数显式收窄，1 基口径） —— *)
_udInLen   := LEN(sIn);                            // 输入字符数 / Input length
_udMarkLen := LEN(sMark);                          // 标记字符数 / Mark length

(* —— 段 4：未超长：原样返回（早退，避免任何改写） —— *)
IF _udInLen <= UINT_TO_UDINT(uiMaxLen) THEN
    sOut       := sIn;                             // 原样返回 / Return as-is
    uiOutLen   := UDINT_TO_UINT(_udInLen);         // 实际长度 / Actual length
    bTruncated := FALSE;                           // 未截断 / Not truncated
    IF eErrCode <> E_DL_StrTruncErr.eClampLen THEN
        eErrCode := E_DL_StrTruncErr.eOk;          // 保留钳位码优先 / Keep clamp code if present
    END_IF
    FC_DL_StringTruncEllipsis := TRUE;             // 结果可信 / Result trustworthy
    RETURN;
END_IF

(* —— 段 5：标记余量判定（标记占满目标长度 → 退化为纯截断） —— *)
IF _udMarkLen >= UINT_TO_UDINT(uiMaxLen) THEN
    _udCopy := UINT_TO_UDINT(uiMaxLen);            // 全部长度用于正文 / All length spent on text
    sOut    := MID(sIn, _udCopy, DL_STE_START);    // 纯截断，无标记 / Plain truncation without mark
    bTruncated := TRUE;
    eErrCode := E_DL_StrTruncErr.eTruncNoMark;     // 信息级：无标记余量 / Info: no room for mark
ELSE
    _udKeep := UINT_TO_UDINT(uiMaxLen) - _udMarkLen;   // 正文保留数 = 目标 - 标记 / Text kept = target - mark
    IF _udKeep < DL_STE_START THEN
        _udKeep := DL_STE_START;                   // 起算位置下限保护（>=1） / Start position lower bound
    END_IF
    sOut    := CONCAT(MID(sIn, _udKeep, DL_STE_START), sMark);  // 正文前缀 + 标记 / Text prefix plus mark
    bTruncated := TRUE;
    eErrCode := E_DL_StrTruncErr.eOk;              // 信息级成功 / Info success
END_IF

(* —— 段 6：结果复检（长度不得超过目标；超限回哨兵） —— *)
uiOutLen := UDINT_TO_UINT(LEN(sOut));              // 实测结果长度 / Measured result length
IF uiOutLen > uiMaxLen THEN
    sOut     := '';                                // 超限回哨兵 / Over-limit to sentinel
    uiOutLen := 0;
    eErrCode := E_DL_StrTruncErr.eInvalidParam;    // 故障级码 / Fault-level code
    RETURN;                                        // 返回 FALSE 保持 / Keep return FALSE
END_IF

FC_DL_StringTruncEllipsis := TRUE;                 // 截断有效 / Truncation valid

END_FUNCTION

(* ---- FC_DL_SurfaceConvectionCalc.st ---- *)
(*
  Component : FC_DL_SurfaceConvectionCalc
  Category  : DL_Base
  Function  : 表面换热系数：自然对流（垂直/水平）与强制对流分式选取
  Complexity: C2
  开源溯源 : DLF 内部原创（R94 族模板派生）；参考语义来源见 SOURCE_HUNTING_MATRIX.md
  规则遵从 : R1-R16
  契约     : 输入 eMode 对流模式枚举、rDeltaTK 表面与环境的温差（取绝对值参与公式） [K]、
             rCharLenM 特征尺寸（垂直取高、水平取宽） [m]、rVelMs 风速（强制模式用） [m/s]；
             输出 rHWm2K 表面换热系数 [W/(m2·K)]、rModeEcho 实际使用模式、
             xValid 有效标志、nFaultCode 故障码。
  边界     : 自然对流派生式 h = 1.42×(ΔT/L)^0.25（垂直）/ 1.32×(ΔT/L)^0.25（水平），
             强制对流简式 h = 10.45×v^0.8；四次方根与 0.8 次幂一律用 EXP(k×LN(x)) 实现，
             禁用 EXPT 等方言算子；ΔT 与 L 须 >0、v 须 >0（强制模式）。
  码位     : 9801 输入非有限（故障级）；9802 特征尺寸或温差越域（故障级）；9803 模式未知（故障级）。
*)
TYPE E_DL_ConvMode :
(
    eNatVertical   := 0,    // 自然对流-垂直面 EN: natural convection on a vertical surface
    eNatHorizontal := 1,    // 自然对流-水平面 EN: natural convection on a horizontal surface
    eForced        := 2     // 强制对流 EN: forced convection
);
END_TYPE

FUNCTION FC_DL_SurfaceConvectionCalc : BOOL
VAR_INPUT
    eMode     : E_DL_ConvMode;   // 对流模式 [-] EN: the convection mode
    rDeltaTK  : LREAL := 30.0;   // 表面与环境温差（取绝对值） [K] EN: the surface to ambient temperature difference taken as a magnitude
    rCharLenM : LREAL := 1.0;    // 特征尺寸 [m] EN: the characteristic length
    rVelMs    : LREAL := 1.0;    // 风速（强制模式） [m/s] EN: the air velocity used in the forced mode
END_VAR
VAR_OUTPUT
    rHWm2K   : LREAL;            // 表面换热系数 [W/(m2·K)] EN: the surface heat transfer coefficient
    rModeEcho: INT;              // 实际使用模式的枚举值 EN: the enumeration value of the mode in use
    xValid   : BOOL;             // 输出可信标志 EN: the outputs are valid
    nFaultCode: INT;             // 0=无故障 9801=输入非有限 9802=尺寸或温差越域 9803=模式未知 EN: zero none, 9801 non finite, 9802 length or difference out of range, 9803 unknown mode
END_VAR
VAR
    xFinAll : BOOL;              // 三个浮点入参有限 EN: the three floating inputs are finite
    rRatio  : LREAL;             // ΔT/L 比 [-] EN: the ratio of the difference to the length
    rPow    : LREAL;             // 幂运算中间值 [-] EN: the interim power value
    rH      : LREAL;             // 换热系数中间值 [W/(m2·K)] EN: the interim coefficient
END_VAR
VAR CONSTANT
    DL_SCV_Z      : LREAL := 0.0;      // 浮点零常量 EN: the floating point zero constant
    DL_SCV_KV     : LREAL := 1.42;     // 垂直自然对流系数 EN: the vertical natural convection factor
    DL_SCV_KH     : LREAL := 1.32;     // 水平自然对流系数 EN: the horizontal natural convection factor
    DL_SCV_KF     : LREAL := 10.45;    // 强制对流系数 EN: the forced convection factor
    DL_SCV_E_NAT  : LREAL := 0.25;     // 自然对流指数 [-] EN: the natural convection exponent
    DL_SCV_E_FRC  : LREAL := 0.8;      // 强制对流指数 [-] EN: the forced convection exponent
    DL_SCV_MIN    : LREAL := 1.0E-6;   // 尺寸与温差的下限 EN: the lower bound of the length and the difference
    DL_SCV_C_BAD  : INT := 9801;       // 输入非有限 EN: a non finite input
    DL_SCV_C_RANG : INT := 9802;       // 尺寸或温差越域 EN: the length or the difference is out of range
    DL_SCV_C_MODE : INT := 9803;       // 模式未知 EN: the mode is unknown
END_VAR

// 段1｜出口预置
FC_DL_SurfaceConvectionCalc := FALSE;   // 返回值预置假 EN: preset the return value to false
rHWm2K := DL_SCV_Z;                     // 换热系数预置零 [W/(m2·K)] EN: preset the coefficient to zero
rModeEcho := 0;                         // 模式回显预置零 EN: preset the mode echo to zero
xValid := FALSE;                        // 有效标志预置假 EN: preset the validity flag to false
nFaultCode := 0;                        // 故障码预置零 EN: preset the fault code to zero

// 段2｜非有限闸：三浮点入参全列（强制模式的风速亦在闸内）
xFinAll := (rDeltaTK = rDeltaTK) AND ((rDeltaTK - rDeltaTK) = DL_SCV_Z)
        AND (rCharLenM = rCharLenM) AND ((rCharLenM - rCharLenM) = DL_SCV_Z)
        AND (rVelMs = rVelMs) AND ((rVelMs - rVelMs) = DL_SCV_Z);   // 三输入有限性 EN: the finiteness of all three inputs
IF NOT xFinAll THEN                                                  // 非有限出口 EN: leave early on a non finite input
    nFaultCode := DL_SCV_C_BAD;                                      // 非有限码 EN: the non finite code
    RETURN;                                                          // 早退 EN: return early
END_IF

// 段3｜域闸：特征尺寸为正、温差取绝对值后须为正（零温差无对流）
IF (rCharLenM < DL_SCV_MIN) OR (ABS(rDeltaTK) < DL_SCV_MIN) THEN      // 尺寸与温差闸 EN: the length and difference gate
    nFaultCode := DL_SCV_C_RANG;                                     // 越域码 EN: the out of range code
    RETURN;                                                          // 早退 EN: return early
END_IF

// 段4｜模式分派：ENUM + CASE 且 ELSE 兜底
rRatio := ABS(rDeltaTK) / rCharLenM;                                 // ΔT/L，分母已证正 [-] EN: the ratio, the divisor is proven positive
CASE eMode OF
    E_DL_ConvMode.eNatVertical:
        rPow := EXP(DL_SCV_E_NAT * LN(rRatio));                      // (ΔT/L)^0.25 EN: the quarter power of the ratio
        rH := DL_SCV_KV * rPow;                                      // 垂直面自然对流 [W/(m2·K)] EN: the vertical natural convection
        rModeEcho := 0;                                              // 模式回显 EN: the mode echo
    E_DL_ConvMode.eNatHorizontal:
        rPow := EXP(DL_SCV_E_NAT * LN(rRatio));                      // (ΔT/L)^0.25 EN: the quarter power of the ratio
        rH := DL_SCV_KH * rPow;                                      // 水平面自然对流 [W/(m2·K)] EN: the horizontal natural convection
        rModeEcho := 1;                                              // 模式回显 EN: the mode echo
    E_DL_ConvMode.eForced:
        IF rVelMs < DL_SCV_MIN THEN                                  // 强制模式需有效风速 EN: the forced mode needs a usable velocity
            nFaultCode := DL_SCV_C_RANG;                             // 风速越域码 EN: the velocity code
            RETURN;                                                  // 早退 EN: return early
        END_IF
        rPow := EXP(DL_SCV_E_FRC * LN(rVelMs));                      // v^0.8 EN: the point eight power of the velocity
        rH := DL_SCV_KF * rPow;                                      // 强制对流 [W/(m2·K)] EN: the forced convection
        rModeEcho := 2;                                              // 模式回显 EN: the mode echo
ELSE
    nFaultCode := DL_SCV_C_MODE;                                     // 未知模式码 EN: the unknown mode code
    RETURN;                                                          // 早退 EN: return early
END_CASE

// 段5｜结果复检与出口
IF (rH <> rH) OR (rH <= DL_SCV_Z) THEN                               // 复检：非有限或非正 EN: recheck for a non finite or non positive value
    nFaultCode := DL_SCV_C_RANG;                                     // 复检失败码 EN: the recheck failure code
    RETURN;                                                          // 早退，出口保持零哨兵 EN: return early with the zero sentinels
END_IF
rHWm2K := rH;                                                        // 换热系数出口 [W/(m2·K)] EN: the coefficient output
xValid := TRUE;                                                      // 结果可信 EN: the results are valid
FC_DL_SurfaceConvectionCalc := TRUE;                                 // 返回真 EN: return true
END_FUNCTION

(* ---- FC_DL_TempDiffUnitConvert.st ---- *)
(*
  FC_DL_TempDiffUnitConvert —— 温差换算 K 与摄氏差值与华氏差值，无偏移项
  分类：DL_Base | 复杂度：1 | 轮次：R86
  开源溯源：道莅原创（clean-room 自研，纯 IEC 61131-3 通用算法），无外部代码引用
  许可证：MIT
  职责：温差（不是温度点！）折算到基准单位 K：开尔文差与摄氏差等价（1:1），
        华氏差 × 5/9。**本件不含 273.15 偏移项**——偏移只属于温度点换算，误用会引入系统偏差。
  契约：fIn 输入温差 [源单位]，eUnit 源单位枚举；fOut 折算结果 [K]；返回 TRUE 表示 fOut 可信。
  边界：① 显式声明无偏移项（分工口径）；② 未知枚举 / 非有限输入 → FALSE + 0.0 哨兵；
        ③ 乘 0.5555555555555556 代替除法，零全局、零物理地址、零库件依赖。
*)

(*-----------------------------------------------------------------------------
 * 枚举: E_DL_TdUnit（温差单位，归属本文件，全库唯一定义）
 *----------------------------------------------------------------------------*)
TYPE E_DL_TdUnit :
(
    eKelvin   := 0,    // 开尔文差值（基准单位） [K] / Kelvin difference, the base unit
    eCelsius  := 1,    // 摄氏差值（与开尔文差 1:1） [K] / Celsius difference, identical to kelvin difference
    eFahrenheit := 2   // 华氏差值（× 5/9） [K] / Fahrenheit difference, scaled by five ninths
);
END_TYPE

FUNCTION FC_DL_TempDiffUnitConvert : BOOL
VAR_INPUT
    fIn   : LREAL := 0.0;              // 输入温差 [源单位] / The input temperature difference
    eUnit : E_DL_TdUnit;               // 源单位枚举 [—] / The source unit enumeration
END_VAR
VAR_OUTPUT
    fOut : LREAL;                      // 折算结果 [K] / The converted difference in kelvin
END_VAR
VAR CONSTANT
    DL_TD_ONE  : LREAL := 1.0;         // 摄氏差折开尔文差的系数（1:1） [-] / Celsius difference to kelvin difference
    DL_TD_FIVE : LREAL := 0.5555555555555556; // 5/9 常数（华氏差折开尔文差） [-] / Five ninths constant
    DL_TD_INF  : LREAL := 1.0E30;      // 非有限 / 越界判据上限 [-] / The magnitude gate
    DL_TD_Z    : LREAL := 0.0;         // 浮点零常量 [K] / The floating point zero constant
END_VAR

FC_DL_TempDiffUnitConvert := FALSE;                       // 返回值预置假 / preset the return false
fOut := DL_TD_Z;                                          // 输出预置零哨兵 [K] / preset the zero sentinel
IF (fIn <> fIn) OR (ABS(fIn) > DL_TD_INF) THEN            // 自反判 NaN 或越限判 Inf / NaN or Inf
    fOut := DL_TD_Z;                                      // 非有限值输出零哨兵 [K] / zero the non finite input
ELSE
    CASE eUnit OF
        E_DL_TdUnit.eKelvin:                              // 基准单位直通 / the base unit passes through
            fOut := fIn;                                  // 直通不换算 [K] / pass through unchanged
            FC_DL_TempDiffUnitConvert := TRUE;            // 结果可信 / the result is valid
        E_DL_TdUnit.eCelsius:                             // 摄氏差与开尔文差等价 / Celsius difference is one to one
            fOut := fIn * DL_TD_ONE;                      // 乘 1.0，无偏移项 [K] / multiply by one, no offset
            FC_DL_TempDiffUnitConvert := TRUE;            // 结果可信 / the result is valid
        E_DL_TdUnit.eFahrenheit:                          // 华氏差折开尔文差 / Fahrenheit difference to kelvin
            fOut := fIn * DL_TD_FIVE;                     // 乘 5/9，无偏移项 [K] / multiply by five ninths, no offset
            FC_DL_TempDiffUnitConvert := TRUE;            // 结果可信 / the result is valid
    ELSE
        fOut := DL_TD_Z;                                  // 未知枚举输出零哨兵 [K] / zero sentinel on an unknown unit
        FC_DL_TempDiffUnitConvert := FALSE;               // 未知枚举不可信 / an unknown unit is not valid
    END_CASE
END_IF
END_FUNCTION

(* ---- FC_DL_VoltageUnitConvert.st ---- *)
(*
  FC_DL_VoltageUnitConvert —— 电压换算 V/mV/kV
  分类：DL_Base | 复杂度：1 | 轮次：R86
  开源溯源：道莅原创（clean-room 自研，纯 IEC 61131-3 通用算法），无外部代码引用
  许可证：MIT
  职责：把电压统一折算到基准单位 V：V 直通、mV 乘 0.001、kV 乘 1000。
  契约：fIn 输入值 [源单位]，eUnit 源单位枚举；fOut 折算结果 [V]；返回 TRUE 表示 fOut 可信。
  边界：未知枚举 / 非有限输入 → 返回 FALSE，fOut 给 0.0 哨兵；无除法，零全局、零物理地址、零库件依赖。
*)

(*-----------------------------------------------------------------------------
 * 枚举: E_DL_VoltUnit（电压单位，归属本文件，全库唯一定义）
 *----------------------------------------------------------------------------*)
TYPE E_DL_VoltUnit :
(
    eVolt     := 0,    // 伏特（基准单位） [V] / Volt, the base unit
    eMilliV   := 1,    // 毫伏 [mV] / Millivolt
    eKiloV    := 2     // 千伏 [kV] / Kilovolt
);
END_TYPE

FUNCTION FC_DL_VoltageUnitConvert : BOOL
VAR_INPUT
    fIn   : LREAL := 0.0;              // 输入值 [源单位] / The input value in the source unit
    eUnit : E_DL_VoltUnit;             // 源单位枚举 [—] / The source unit enumeration
END_VAR
VAR_OUTPUT
    fOut : LREAL;                      // 折算结果 [V] / The converted value in the base unit
END_VAR
VAR CONSTANT
    DL_VT_MV  : LREAL := 0.001;        // 1 mV 折 V 的系数 [-] / millivolt to volt
    DL_VT_KV  : LREAL := 1000.0;       // 1 kV 折 V 的系数 [-] / kilovolt to volt
    DL_VT_INF : LREAL := 1.0E30;       // 非有限 / 越界判据上限 [-] / The magnitude gate
    DL_VT_Z   : LREAL := 0.0;          // 浮点零常量 [V] / The floating point zero constant
END_VAR

FC_DL_VoltageUnitConvert := FALSE;                        // 返回值预置假 / preset the return false
fOut := DL_VT_Z;                                          // 输出预置零哨兵 [V] / preset the zero sentinel
IF (fIn <> fIn) OR (ABS(fIn) > DL_VT_INF) THEN            // 自反判 NaN 或越限判 Inf / NaN or Inf
    fOut := DL_VT_Z;                                      // 非有限值输出零哨兵 [V] / zero the non finite input
ELSE
    CASE eUnit OF
        E_DL_VoltUnit.eVolt:                              // 基准单位直通 / the base unit passes through
            fOut := fIn;                                  // 直通不换算 [V] / pass through unchanged
            FC_DL_VoltageUnitConvert := TRUE;             // 结果可信 / the result is valid
        E_DL_VoltUnit.eMilliV:                            // 毫伏折伏 / millivolt to volt
            fOut := fIn * DL_VT_MV;                       // 乘 0.001 [V] / multiply by the factor
            FC_DL_VoltageUnitConvert := TRUE;             // 结果可信 / the result is valid
        E_DL_VoltUnit.eKiloV:                             // 千伏折伏 / kilovolt to volt
            fOut := fIn * DL_VT_KV;                       // 乘 1000 [V] / multiply by the factor
            FC_DL_VoltageUnitConvert := TRUE;             // 结果可信 / the result is valid
    ELSE
        fOut := DL_VT_Z;                                  // 未知枚举输出零哨兵 [V] / zero sentinel on an unknown unit
        FC_DL_VoltageUnitConvert := FALSE;                // 未知枚举不可信 / an unknown unit is not valid
    END_CASE
END_IF
END_FUNCTION

(* ---- FC_DL_ArrCopySeg.st ---- *)
// ==============================================================================
// 组件名 Component  : FC_DL_ArrCopySeg
// 分类   Category   : DL_Base
// 前缀   Naming     : FC_DL_ ｜ b/n/i/f 类型前缀制（R265）
// 版本   Version    : 1.0.0
// 复杂度 Complexity  : 低
// 功能   Purpose    : 定长 LREAL 数组段拷贝：把源数组 [iSrcFrom ..] 起的
//                      nCnt 个元素拷到目标数组 [iDstFrom ..] 起；nCnt <= 0
//                      零拷贝合法；源 / 目标越界自动截断 nCnt，bTrunc 置位
//                      报告截断，nCopied 反映实际拷贝数（bValid 保持 TRUE）。
//                      供缓冲搬运 / 窗段平移 / 队列重组类调用方使用。
// 开源溯源 Origin    : 西门子 LGF 分类语义借鉴，clean-room 重写（LGF
//                      Data Handling「定长缓冲搬运（无动态内存）」分类学
//                      口径借鉴，只借骨不抄肉，实现零代码复制）
// 许可证 License    : MIT
// 参考   Reference  : IEC 61131-3:2013 §6.6.4 FOR 遍历与数组语义
// 平台   Platform   : 纯 IEC 61131-3（FOR / 数组 / 比较），三平台通用
// 依赖   Depends    : 无（零委托、零库件）
// 分工声明 Split     : FC_DL_ArrFillEx（常数填充）与本件互引；本件为数组段
//                      搬运（源是数组），彼件为常数填充（源是标量），语义
//                      正交（R216）。与 FC_DL_ArraySliceCopy（DL_MathData）
//                      分工：彼件从下标 0 起承接且对越域判故障早退，本件
//                      支持任意目标起点且对越界截断续行（bTrunc 报告），
//                      口径不同勿混用（R216）。
// 归属 Ownership     : 本件无 TYPE 声明；全部引脚为 IEC 标准原生类型。
// ------------------------------------------------------------------
// 边界 Boundary     :
//   一 零拷贝闸：nCnt <= 0 → nCopied = 0、bValid = TRUE、数组零写回
//      （合法语义不是故障）；
//   二 截断闸（逐项点名，R272）：iSrcFrom < 0 / iDstFrom < 0 钳 0 置
//      bTrunc；nCnt 超过源余量（255 - iSrcC）或目标余量（255 - iDstC）
//      时截到较小余量并置 bTrunc；起点越出容量（> 255）时余量为负、
//      nUse <= 0 → 零拷贝 + bTrunc（bValid 保持 TRUE，截断是信息级）；
//   三 重叠自检（中转缓冲两段式）：先把源段整段读入局部 afStaging，再
//      整段写回目标——arrSrc 与 arrDst 为同一数组且区间重叠的别名调用
//      也不产生撕裂 / 串写（快照语义，真实可达：调用方传同一数组做段
//      平移）；此为机制性防重叠，非永假防御；
//   四 拷贝序：读侧 / 写侧循环上界由段 2 截断闸证明 <= 255，下标越界
//      不可达；
//   五 纯函数：无记忆量、无定时器、无边沿实例，每调用重算；
//   六 无除法、无浮点比较；无全局、无外部变量、无物理地址。
// 错误码 Codes      :
//   16#0001_0745【信息级】段越界自动截断（起点钳位或 nCnt 截到余量，
//                bTrunc = TRUE、bValid = TRUE、nCopied 反映实际拷贝数）
//   注：本件引脚契约按任务定稿无独立 eErr 出口，截断语义经 bTrunc /
//   nCopied 双通道表达；零拷贝与截断为零的出口同形（bTrunc 区分），
//   不另设码（R90 反证句）。
// 验收 Acceptance   :
//   算法已证（脚本）：未跑 ｜ 编译器已证（三平台）：未跑
//   V1 源 [1..5]、iSrcFrom = 1、iDstFrom = 10、nCnt = 3 → 目标槽 10..12
//      为 [2,3,4]、nCopied = 3、bTrunc = FALSE
//   V2 nCnt = 0 / 负数 → nCopied = 0、bValid = TRUE、bTrunc = FALSE
//   V3 iSrcFrom = 250、nCnt = 10 → 截到 6、bTrunc = TRUE
//   V4 iSrcFrom = -3 → 钳 0 续拷、bTrunc = TRUE
//   V5 iDstFrom = 300 → nCopied = 0、bTrunc = TRUE
//   V6 别名调用：同一数组段平移 → 中转缓冲两段式无撕裂（V1 断言不变）
// 修订记录 Revision  :
//   2026-11-22  v1.0.0  R65 首版（批 1 · 序号 4，LGF Data Handling 补口）
// ==============================================================================
FUNCTION FC_DL_ArrCopySeg : BOOL
VAR_IN_OUT
    arrSrc : ARRAY[0..255] OF LREAL; // 源数组 [工程单位]，允许与目标同数组（别名调用走中转缓冲）/ the source array, may alias the target
    arrDst : ARRAY[0..255] OF LREAL; // 目标数组 [工程单位]，从 iDstFrom 起承接 / the target array receiving from iDstFrom
END_VAR
VAR_INPUT
    iSrcFrom : INT := 0;         // 源段起点 [下标]，负值钳 0 / the source start index, negative clamped
    iDstFrom : INT := 0;         // 目标段起点 [下标]，负值钳 0 / the target start index, negative clamped
    nCnt     : INT := 0;         // 请求拷贝数 [个]，<= 0 零拷贝合法 / the requested count, zero or less is a legal no op
END_VAR
VAR_OUTPUT
    nCopied : INT;               // 实际拷贝数 [个] / the actually copied count
    bValid  : BOOL;              // 结果可用 [-]，本件恒 TRUE（截断为信息级）/ the validity flag, always true here
    bTrunc  : BOOL;              // 截断报告 [-]，TRUE = 发生钳位或截断 / the truncation flag
END_VAR
VAR
    iSrcC     : INT;             // 钳位后的源起点 [下标] / the clamped source start
    iDstC     : INT;             // 钳位后的目标起点 [下标] / the clamped target start
    nAvail    : INT;             // 源 / 目标余量的较小值 [个] / the smaller of the two remainders
    nUse      : INT;             // 实际拷贝数暂存 [个] / the staged copy count
    k         : INT;             // 遍历索引 [下标] / the traversal index
    afStaging : ARRAY[0..255] OF LREAL; // 中转缓冲 [工程单位]，两段式防重叠撕裂 / the staging buffer for the overlap safe two stage copy
END_VAR
VAR CONSTANT
    DL_ACP_NMAX : INT := 255;    // 数组容量上界 [个]，与数组容量一致 / the capacity aligned with the array
    DL_ACP_ZERO : INT := 0;      // 整型零常量 [个] / the integer zero constant
END_VAR

// 段 1｜返回值与全部出口预置 + 中转缓冲清零（R45 四段式第一段）/ segment 1, the preset and the staging clear
FC_DL_ArrCopySeg := FALSE;       // 返回值预置假 / preset the return false
nCopied := DL_ACP_ZERO;          // 拷贝数预置零 [个] / preset the copied count zero
bValid  := TRUE;                 // 有效标志预置真（截断为信息级口径）/ preset valid
bTrunc  := FALSE;                // 截断标志预置假 / preset the truncation flag false
FOR k := DL_ACP_ZERO TO DL_ACP_NMAX DO // 中转缓冲全量预清零 / preset the staging buffer zero
    afStaging[k] := 0.0;         // 缓冲槽位显式清零 [工程单位] / clear the staging slot explicitly
END_FOR

// 段 2｜截断闸第一段：负起点钳 0 置 bTrunc（边界二，逐项点名）/ segment 2, the clamp of negative starts
iSrcC := iSrcFrom;               // 源起点接管 / take the source start
iDstC := iDstFrom;               // 目标起点接管 / take the target start
IF iSrcC < DL_ACP_ZERO THEN      // 源起点下越界 / the source start below the domain
    iSrcC := DL_ACP_ZERO;        // 钳 0 续拷（信息级 0745）/ clamp to zero and keep copying
    bTrunc := TRUE;              // 置截断报告 / raise the truncation flag
END_IF
IF iDstC < DL_ACP_ZERO THEN      // 目标起点下越界 / the target start below the domain
    iDstC := DL_ACP_ZERO;        // 钳 0 续拷（信息级 0745）/ clamp to zero and keep copying
    bTrunc := TRUE;              // 置截断报告 / raise the truncation flag
END_IF

// 段 3｜零拷贝闸（边界一：nCnt <= 0 合法，数组零写回）/ segment 3, the zero copy gate
IF nCnt <= DL_ACP_ZERO THEN      // 请求拷贝数非正 / the requested count non positive
    nCopied := DL_ACP_ZERO;      // 零拷贝 [个] / a zero copy
    FC_DL_ArrCopySeg := TRUE;    // 合法返回 / return success
    RETURN;                      // 早退，数组零写回 / early return untouched
END_IF

// 段 4｜截断闸第二段：nCnt 截到源 / 目标余量较小值（边界二）/ segment 4, the truncation to the smaller remainder
nAvail := DL_ACP_NMAX - iSrcC;   // 源余量 [个] / the source remainder
IF (DL_ACP_NMAX - iDstC) < nAvail THEN // 目标余量更小 / the target remainder smaller
    nAvail := DL_ACP_NMAX - iDstC; // 取目标余量 [个] / take the target remainder
END_IF
nUse := nCnt;                    // 请求拷贝数接管 [个] / take the requested count
IF iSrcC > DL_ACP_NMAX THEN      // 源起点越出容量 / the source start beyond the capacity
    bTrunc := TRUE;              // 置截断报告（余量为负，落零拷贝）/ raise the truncation flag
END_IF
IF iDstC > DL_ACP_NMAX THEN      // 目标起点越出容量 / the target start beyond the capacity
    bTrunc := TRUE;              // 置截断报告 / raise the truncation flag
END_IF
IF nUse > nAvail THEN            // 请求量超余量 / the request above the remainder
    nUse := nAvail;              // 截到余量（信息级 0745）/ truncate to the remainder
    bTrunc := TRUE;              // 置截断报告 / raise the truncation flag
END_IF
IF nUse <= DL_ACP_ZERO THEN      // 截断后为非正（起点越出容量路径）/ the truncated count non positive
    nCopied := DL_ACP_ZERO;      // 零拷贝 [个] / a zero copy
    FC_DL_ArrCopySeg := TRUE;    // 合法返回 / return success
    RETURN;                      // 早退，数组零写回 / early return untouched
END_IF

// 段 5｜中转缓冲承接源段（边界三：两段式第一段，读侧快照）/ segment 5, the staging takes the source segment
FOR k := DL_ACP_ZERO TO nUse - 1 DO // 有界遍历（上界 = nUse - 1 <= 254 已证）/ the bounded traversal
    afStaging[k] := arrSrc[iSrcC + k]; // 源段读入缓冲 [工程单位]（下标 <= 255 已证）/ read the source into the staging
END_FOR

// 段 6｜缓冲写回目标段（边界三：两段式第二段，写侧顺序落位）/ segment 6, the staging lands on the target
FOR k := DL_ACP_ZERO TO nUse - 1 DO // 有界遍历（上界同段 5 已证）/ the bounded traversal
    arrDst[iDstC + k] := afStaging[k]; // 缓冲整段写回目标 [工程单位]（下标 <= 255 已证）/ land the staging onto the target
END_FOR

// 段 7｜统一出口 / segment 7, the unified outlet
nCopied := nUse;                 // 实拷贝数出口 [个] / the copied count outlet
FC_DL_ArrCopySeg := TRUE;        // 返回成功 / return success
END_FUNCTION

(* ---- FC_DL_ArrFillEx.st ---- *)
// ==============================================================================
// 组件名 Component  : FC_DL_ArrFillEx
// 分类   Category   : DL_Base
// 前缀   Naming     : FC_DL_ ｜ b/n/i/f 类型前缀制（R265）
// 版本   Version    : 1.0.0
// 复杂度 Complexity  : 低
// 功能   Purpose    : 定长 LREAL 数组区间填充：把 [iFrom, iTo] 闭区间各槽位
//                      写为 fVal；区间越界自动钳位（iFrom < 0 钳 0、
//                      iTo > 255 钳 255），iFrom > iTo 零填充合法返回；
//                      bFillNaN = FALSE 且 fVal 非有限时拒绝填充
//                      （bValid = FALSE，数组零写回）。供清屏 / 预置 /
//                      坏点填充类调用方使用。
// 开源溯源 Origin    : 西门子 LGF 分类语义借鉴，clean-room 重写（LGF
//                      Data Handling「定长缓冲批量写」分类学口径借鉴，只借
//                      骨不抄肉，实现零代码复制）
// 许可证 License    : MIT
// 参考   Reference  : IEC 61131-3:2013 §6.6.4 FOR 遍历与数组语义
// 平台   Platform   : 纯 IEC 61131-3（FOR / 数组 / 比较），三平台通用
// 依赖   Depends    : 无（零委托、零库件）
// 分工声明 Split     : FC_DL_ArrCopySeg（段拷贝）与本件互引；本件为常数填充
//                      （源是标量），彼件为数组段搬运（源是数组），语义正交
//                      （R216）。
// 归属 Ownership     : 本件无 TYPE 声明；全部引脚为 IEC 标准原生类型。
// ------------------------------------------------------------------
// 边界 Boundary     :
//   一 区间钳位闸（逐项点名，R272）：iFrom < 0 钳 0、iTo > 255 钳 255，
//      钳位后照常填充（信息级语义，bValid 保持 TRUE）；iFrom / iTo 反向
//      （含钳位后反向）→ 零填充合法返回（nFilled = 0、bValid = TRUE）；
//   二 非有限闸：fVal 为 NaN（自反判 x <> x）或 ±Inf（差值自反判
//      (x - x) <> (x - x)）且 bFillNaN = FALSE → bValid = FALSE、
//      nFilled = 0、数组零写回早退（R272 非有限防护）；bFillNaN = TRUE
//      时允许显式填充 NaN / Inf（调用方自担，bValid 保持 TRUE）；
//   三 填充序：FOR 闭区间顺序写，上界 iToC <= 255、下界 iFromC >= 0 已证
//      （钳位闸证明），下标越界不可达；
//   四 纯函数：无记忆量、无定时器、无边沿实例，每调用重算；
//   五 无除法；无全局、无外部变量、无物理地址。
// 错误码 Codes      :
//   16#0001_0743【信息级】区间越界已钳位续填（iFrom 钳 0 / iTo 钳 255，
//                bValid = TRUE，nFilled 反映实际填充数）
//   16#0001_0744【故障级】fVal 非有限且 bFillNaN = FALSE，拒绝填充
//                （bValid = FALSE、nFilled = 0、数组零写回）
//   注：本件引脚契约按任务定稿无独立 eErr 出口，上述码位为文档级语义，
//   经 bValid / nFilled 通道表达；钳位续填与正常填充出口同形（仅区间
//   收窄），无独立输出通道可承载，不另设出口位（R90 反证句）。
// 验收 Acceptance   :
//   算法已证（脚本）：未跑 ｜ 编译器已证（三平台）：未跑
//   V1 iFrom = 10、iTo = 20、fVal = 5.0 → 槽位 10..20 全为 5.0、nFilled = 11
//   V2 iFrom = -5 → 钳 0 续填；iTo = 300 → 钳 255 续填
//   V3 iFrom > iTo → nFilled = 0、bValid = TRUE、数组原样
//   V4 fVal = NaN、bFillNaN = FALSE → bValid = FALSE、零写回
//   V5 fVal = NaN、bFillNaN = TRUE → 填入 NaN、bValid = TRUE
// 修订记录 Revision  :
//   2026-11-22  v1.0.0  R65 首版（批 1 · 序号 3，LGF Data Handling 补口）
// ==============================================================================
FUNCTION FC_DL_ArrFillEx : BOOL
VAR_IN_OUT
    arrDst : ARRAY[0..255] OF LREAL; // 目标数组 [工程单位]，闭区间填充 / the target array filled over the closed range
END_VAR
VAR_INPUT
    iFrom    : INT;              // 填充起点 [下标]，闭区间含端点 / the fill start index, inclusive
    iTo      : INT;              // 填充终点 [下标]，闭区间含端点 / the fill end index, inclusive
    fVal     : LREAL;            // 填充值 [工程单位] / the fill value
    bFillNaN : BOOL := FALSE;    // 允许非有限填充开关 [-]，TRUE 时允许填 NaN / Inf / the non finite fill switch
END_VAR
VAR_OUTPUT
    nFilled : INT;               // 实际填充槽位数 [个] / the actually filled slot count
    bValid  : BOOL;              // 结果可用 [-]，拒绝填充为 FALSE / the result usable flag
END_VAR
VAR
    iFromC     : INT;            // 钳位后的填充起点 [下标] / the clamped fill start
    iToC       : INT;            // 钳位后的填充终点 [下标] / the clamped fill end
    k          : INT;            // 遍历索引 [下标] / the traversal index
    xNonFinite : BOOL;           // fVal 非有限标志 [-] / the non finite flag of fVal
END_VAR
VAR CONSTANT
    DL_AFE_NMAX : INT := 255;    // 数组容量上界 [个]，与数组容量一致 / the capacity aligned with the array
    DL_AFE_ZERO : INT := 0;      // 整型零常量 [个] / the integer zero constant
END_VAR

// 段 1｜返回值与全部出口预置（R45 四段式第一段）/ segment 1, the preset of the return and all outlets
FC_DL_ArrFillEx := FALSE;        // 返回值预置假 / preset the return false
nFilled := DL_AFE_ZERO;          // 填充数预置零 [个] / preset the filled count zero
bValid  := TRUE;                 // 有效标志预置真（零填充合法口径）/ preset valid, a legal zero fill

// 段 2｜区间钳位闸（边界一：iFrom 钳 0 / iTo 钳 255，逐项点名）/ segment 2, the range clamp gate
iFromC := iFrom;                 // 起点接管 / take the start
iToC   := iTo;                   // 终点接管 / take the end
IF iFromC < DL_AFE_ZERO THEN     // 起点下越界 / the start below the domain
    iFromC := DL_AFE_ZERO;       // 钳 0 续填（信息级 0743）/ clamp to zero and keep filling
END_IF
IF iToC > DL_AFE_NMAX THEN       // 终点上越界 / the end above the domain
    iToC := DL_AFE_NMAX;         // 钳 255 续填（信息级 0743）/ clamp to the cap and keep filling
END_IF

// 段 3｜反向区间闸：零填充合法返回（边界一）/ segment 3, the reversed range gate, a legal zero fill
IF iFromC > iToC THEN            // 起点 > 终点（含钳位后反向）/ the start above the end
    nFilled := DL_AFE_ZERO;      // 零填充 [个] / a zero fill
    FC_DL_ArrFillEx := TRUE;     // 合法返回 / return success
    RETURN;                      // 早退，数组零写回 / early return untouched
END_IF

// 段 4｜非有限闸（边界二：NaN 自反判 + Inf 差值自反判，R272）/ segment 4, the non finite gate
xNonFinite := (fVal <> fVal) OR ((fVal - fVal) <> 0.0); // NaN 或 ±Inf / NaN or infinity
IF (NOT bFillNaN) AND xNonFinite THEN // 未允许且非有限 / not allowed and non finite
    bValid  := FALSE;            // 拒绝填充（故障级 0744）/ refuse the fill
    nFilled := DL_AFE_ZERO;      // 填充数归零 [个] / zero the count
    FC_DL_ArrFillEx := FALSE;    // 返回失败 / return failure
    RETURN;                      // 早退，数组零写回 / early return untouched
END_IF

// 段 5｜闭区间顺序填充（边界三：上界已证 <= 255、下界已证 >= 0）/ segment 5, the ordered closed range fill
FOR k := iFromC TO iToC DO       // 有界遍历 / the bounded traversal
    arrDst[k] := fVal;           // 槽位写入 [工程单位] / write the slot
END_FOR

// 段 6｜统一出口 / segment 6, the unified outlet
nFilled := iToC - iFromC + 1;    // 实际填充数 [个] / the actually filled count
FC_DL_ArrFillEx := TRUE;         // 返回成功 / return success
END_FUNCTION

(* ---- FC_DL_BinaryToGray.st ---- *)
(*==============================================================================
 * 组件名称 (Component)  : FC_DL_BinaryToGray
 * 所属子库 (Sublibrary) : DL_Base
 * 当前版本 (Version)    : 1.0.0
 * 兼容性   (Platform)   : CODESYS 3.5 / TwinCAT 3 / 汇川 InoProShop / Machine Expert
 *                         仅用标准 SHL / SHR / XOR / AND，无厂商方言
 * 功能描述 (Function)   : 二进制 → 格雷码纯映射函数，用于"向绝对值编码器写目标位置"
 *                         以及"生成格雷码测试序列验证 FC_DL_GrayToBinary"。
 *                         与 FC_DL_GrayToBinary 严格互逆：GrayToBinary(BinaryToGray(x)) = x
 *                         （x 位于 0..2^w-1 且位宽一致时）。
 *                         输入先掩码再去脏高位；位宽 32 时掩码特判全 1，避免 SHL(1,32)。
 * 算法     (Algorithm)  : G = (B XOR (B >> 1)) AND mask，单表达式实现，禁止 FOR。
 * 开源溯源 (Origin)     : 原创实现。格雷码定义为公开经典算法，掩码与钳位为本库工程加固。
 * 依赖     (Depends)    : 无 DL_ 内部依赖；无标准库功能块依赖
 * 互逆性自检 (Inverse Check): 手册给出的验证用例——对 0..2^w-1 全序列，
 *                         FC_DL_GrayToBinary(FC_DL_BinaryToGray(x, w), w) 必须等于 x。
 * 红线自检 (Redline)    : R1 ✓ 零全局变量表与外部变量引用 ｜ R2 ✓ 零物理 IO 地址直写
 *                         R3 ✓ 纯 IEC 61131-3 ｜ R4 ✓ 位宽钳位 + SHL(1,32) 特判 + 先掩码后异或
 *                         R5 ✓ 全变量中英双语同行注释 ｜ R6 N/A（无状态机）｜ R7 N/A（无实例调用）
 * 修订历史 (Revision)   :
 *   2026-11-14  v1.0.0  首版入库（Phase 1 冷启动 · Level 0 批次）
 *============================================================================*)
FUNCTION FC_DL_BinaryToGray : UDINT
VAR_INPUT
    uBinaryValue : UDINT;         // 二进制原始值，允许带高位脏数据 / Raw binary value, dirty high bits tolerated
    uBitWidth    : USINT := 32;   // 有效位宽 1..32，越界按边界钳位 / Valid bit width 1..32, clamped at the boundaries
END_VAR
VAR_OUTPUT
    bValid       : BOOL;          // 位宽合法标志，FALSE 表示参数越界已钳位 / Width valid flag, FALSE means clamped
    uErrorId     : UDINT;         // 故障码，0 = 无故障 / Error code, 0 = no error
END_VAR
VAR
    uMask        : UDINT;         // 位宽掩码，仅保留有效位 / Bit-width mask keeping valid bits only
    uWidth       : USINT;         // 钳位后的有效位宽 / Clamped effective bit width
    uMaskedValue : UDINT;         // 已剔除脏高位的规范化输入 / Normalized input with dirty high bits removed
END_VAR
VAR CONSTANT
    DL_GRAY_WIDTH_MIN : USINT := 1;    // 最小合法位宽 [bit] / Min legal bit width [bit]
    DL_GRAY_WIDTH_MAX : USINT := 32;   // 最大合法位宽 [bit] / Max legal bit width [bit]
END_VAR

(*------------------------------------------------------------------------------
 * 段 1｜返回值与工作变量预置：任何路径下返回值确定
 *      Initialize return value and working variables for determinism
 *-----------------------------------------------------------------------------*)
FC_DL_BinaryToGray := 16#0000_0000;
bValid             := TRUE;
uErrorId           := 16#0000_0000;
uMask              := 16#0000_0000;
uWidth             := uBitWidth;
uMaskedValue       := 16#0000_0000;

(*------------------------------------------------------------------------------
 * 段 2｜位宽钳位（边界 B1）：钳位 + 告警，但继续计算有效结果
 *      Width clamping: clamp and warn while still producing a valid result
 *-----------------------------------------------------------------------------*)
IF uBitWidth < DL_GRAY_WIDTH_MIN THEN
    uWidth   := DL_GRAY_WIDTH_MIN;
    bValid   := FALSE;
    uErrorId := 16#0001_0001;
ELSIF uBitWidth > DL_GRAY_WIDTH_MAX THEN
    uWidth   := DL_GRAY_WIDTH_MAX;
    bValid   := FALSE;
    uErrorId := 16#0001_0001;
END_IF

(*------------------------------------------------------------------------------
 * 段 3｜掩码构造（边界 B2）：位宽 32 特判全 1，绝不执行 SHL(1,32)
 *      Mask construction: all-ones at width 32, SHL(1,32) is never executed
 *-----------------------------------------------------------------------------*)
IF uWidth >= DL_GRAY_WIDTH_MAX THEN
    uMask := 16#FFFF_FFFF;
ELSE
    uMask := SHL(UDINT#1, USINT_TO_UDINT(uWidth)) - 16#0000_0001;
END_IF

(*------------------------------------------------------------------------------
 * 段 4｜先掩码（边界 B4）：顺序不可交换
 *      Mask first: the order is not interchangeable
 *      若先异或后掩码，脏高位会经右移渗入有效位区间，掩码只能截断结果、
 *      无法还原已被污染的低位，因此必须先规范化输入
 *-----------------------------------------------------------------------------*)
uMaskedValue := uBinaryValue AND uMask;

(*------------------------------------------------------------------------------
 * 段 5｜单表达式转换（边界 B3）：G = (B XOR (B >> 1)) AND mask
 *      Single-expression conversion, no loop by design
 *-----------------------------------------------------------------------------*)
FC_DL_BinaryToGray := (uMaskedValue XOR SHR(uMaskedValue, 1)) AND uMask;
END_FUNCTION

(* ---- FC_DL_BitArrayInsert.st ---- *)
(*==============================================================================
 * 组件名称 (Component)  : FC_DL_BitArrayInsert
 * 所属子库 (Sublibrary) : DL_Base
 * 归属目录 (Directory)  : C:\Library\DL_Base
 * 当前版本 (Version)    : 1.0.0
 * 组件分类 (Category)   : 函数（FUNCTION）· 原子位窗写 · 跨字读改写
 * 兼容性   (Platform)   : CODESYS 3.5 / TwinCAT 3 / 汇川 InoProShop / 施耐德
 *                         Machine Expert；仅用 Standard.library 的 SHL / SHR /
 *                         AND / OR / NOT 与显式类型转换，无厂商位访问方言
 * 功能一句话 (Summary)  : 把 64 位值按「起始位 + 位宽」原子写入 DWORD 数组位流的
 *                         指定窗口，只改窗口内的位，并报出实际改动字数。
 * 功能描述 (Function)   : 与 FC_DL_BitArrayExtract 严格成对：提取件读窗口，
 *                         本件写窗口。窗口跨字时先算出两个字的完整新值，再按
 *                         低字、高字顺序一次性回写，避免半更新撕裂。
 *                         典型现场用途：64 位使能字与报警屏蔽字下发、凸轮表位图
 *                         整段更新、远程 IO 位图按字段改写而不动邻位。
 * 与既有件边界 (Boundary): FC_DL_BitSet 只置单字内单个位；FC_DL_WordBitPack 只把
 *                         多个位段打包进一个 WORD；本件是跨字位流窗口的读改写，
 *                         带改动计数与原子写回语义，三者职责互斥。
 * 副作用声明 (Side effect): 本件是「纯函数语义 + 受控副作用」：无内部状态、同入参
 *                         同结果，但会原地修改形参指向的目标数组。副作用范围仅限
 *                         形参数组的窗口内位，绝不触碰窗口外位，也绝不写数组之外。
 *                         严禁把本件当只读函数使用。
 * 设计要点 (Key notes)  : ① 先算完全部新值再回写，杜绝读一半写一半；
 *                         ② 先比较后计数：值未变的字不计入改动数，也不产生写动作，
 *                           减少下游无谓刷新；
 *                         ③ 宽度 64 走满 1 常量分支，禁止左移 64 位；
 *                         ④ 越界截断后仍写可用位并置 bValid 为假，现场可读可查。
 * 开源溯源 (Origin)     : 来源标签 lgf-bitlogic。LGF 为免费闭源发布的公开函数库
 *                         手册，本件仅借鉴其位逻辑组「打包与提取双向成对」的组织
 *                         方式与「批量位串三口分工」的分类骨架；许可证按其发布方
 *                         条款仅作分类参考，本件零代码行、零注释、零数据结构引用，
 *                         属 clean-room 独立实现，不构成衍生作品。
 * 码位说明 (Codes)      : 本件独占信息级码段 16#0001_0128 到 16#0001_012A，纯函数
 *                         语义无锁存面故不占故障级码；与提取件的 0125 到 0127 相邻
 *                         不重叠，与全库已占码求差为空。
 *                         0128 偏移越界 ｜ 0129 宽度越界 ｜ 012A 跨字截断。
 * 依赖说明 (Depends)    : 无 DL_ 内部依赖；仅 Standard.library 的 SHL / SHR / NOT /
 *                         DWORD_TO_LWORD / LWORD_TO_DWORD / INT_TO_DINT / INT_TO_UDINT。
 * 契约前置条件 (Contract): 函数内无法探测数组实际长度，故「nTargetCount 不得大于
 *                         调用方实际数组长度」由调用方负责，组态时须保证。
 * 红线自检 (Redline)    : 零全局变量表依赖 ｜ 零外部变量声明 ｜ 零物理地址
 *                         纯 IEC 61131-3 ｜ 无除法故无除零面 ｜ 全变量双语同行注释
 *                         状态机 N/A（纯函数）｜ 无定时器实例 ｜ 移位量恒小于 64
 * 修订历史 (Revision)   : 2026-11-15  v1.0.0  首版入库（Round 12 · 跨字位段族）
 *============================================================================*)

(*==============================================================================
 * 读改写示意 (Read modify write)：
 *   目标两字初值 16#FFFF_FFFF 与 16#FFFF_FFFF，起始位 28、位宽 8、写入 16#A5
 *   掩码 16#FF 左移 28 位后覆盖第 1 字的高 4 位与第 2 字的低 4 位
 *   第 1 字新值 16#5FFF_FFFF，第 2 字新值 16#FFFF_FFFA，改动字数 2
 *   窗口外的位一字不动，这是本件与「整字覆盖」最本质的差别
 *============================================================================*)

(*==============================================================================
 * 逐调用推演 (Call trace)：
 *   调用 1  初值全 1、起始 28、位宽 8、写入 16#A5
 *     字数 2，总位数 64；偏移 28 通过；宽度 8 通过；28 加 8 等于 36 不截断
 *     低字下标 1，移位 28，跨字判据成立，高字下标 2
 *     掩码 16#FF，生效值 16#A5，展开后低字得 16#5FFF_FFFF、高字得 16#FFFF_FFFA
 *     两字都与旧值不同，改动计数 2，写回后返回真
 *   调用 2  初值 16#0000_000F、起始 0、位宽 4、写入 16#F
 *     新值与旧值相同，改动计数 0，不发写动作，目标保持原值
 *   调用 3  起始 30、位宽 8、字数 1、写入 16#FF
 *     30 加 8 超过 32，宽度截为 2，事件码 012A，只写最高两位的 16#3
 *============================================================================*)

FUNCTION FC_DL_BitArrayInsert : BOOL
VAR_IN_OUT
    auTarget     : ARRAY[1..8] OF DWORD;  // 被写入的目标位流数组，本函数原地修改窗口内位 [位串] / Target bit stream, window bits modified in place
END_VAR
VAR_INPUT
    uValue       : LWORD;                 // 待写入值，只用低 nWidth 位，超宽位忽略 [位串] / Value to write, only the low window bits are used
    nTargetCount : INT := 1;              // 目标有效字数 [个]，域 1 到 8，越界钳位 / Effective target word count, 1 to 8, clamped
    nOffset      : INT := 0;              // 写入窗口起始位 [bit]，0 起 / Window start bit, zero based
    nWidth       : INT := 8;              // 写入窗口宽度 [bit]，域 1 到 64 / Window width, 1 to 64
END_VAR
VAR_OUTPUT
    nChanged     : INT;                   // 实际发生改动的字数 [个]，值未变的字不计入 / Number of words actually modified
    uApplied     : LWORD;                 // 实际写入的右对齐值，已按宽度截断 [位串] / Value actually applied, width masked
    uMask        : LWORD;                 // 本次生效掩码，右对齐 [位串] / Effective right aligned mask
    nActualW     : INT;                   // 实际生效宽度 [bit] / Effective width after truncation
    uErrorId     : UDINT;                 // 事件码，0 表示无事件 / Event code, zero means none
    bValid       : BOOL;                  // 全合法为真，截断或越界为假 / All inputs legal, false when truncated
END_VAR
VAR
    nTotalBits   : DINT;                  // 目标位流总位数，等于字数乘 32 [bit] / Total bit count of the target stream
    nIdxLo       : INT;                   // 低字下标，1 起 [索引] / Low word index, one based
    nIdxHi       : INT;                   // 高字下标，0 表示不跨字 [索引] / High word index, zero when not straddling
    nShift       : INT;                   // 字内移位量，等于偏移对 32 取模 [bit] / Intra word shift amount
    uWinWide     : LWORD;                 // 已左移到窗口位置的写入值 [位串] / Window value shifted into place
    uMaskWide    : LWORD;                 // 已左移到窗口位置的掩码 [位串] / Window mask shifted into place
    uOldLo       : DWORD;                 // 低字旧值 [位串] / Previous low word
    uOldHi       : DWORD;                 // 高字旧值，不跨字时为 0 [位串] / Previous high word, zero when absent
    uNewLo       : DWORD;                 // 低字新值 [位串] / New low word
    uNewHi       : DWORD;                 // 高字新值，不跨字时为 0 [位串] / New high word, zero when absent
END_VAR
VAR CONSTANT
    DL_MASK64_ALL : LWORD := 16#FFFF_FFFF_FFFF_FFFF;   // 满宽掩码常量，64 宽分支专用 [位串] / All ones mask for the 64 bit branch
    DL_SRC_MAX    : INT := 8;                          // 目标字数上限 [个] / Target word count limit
    DL_BIT_MAX64  : INT := 64;                         // 位窗宽度上限 [bit] / Window width limit
    DL_BIT_MAX32  : INT := 32;                         // 单字位宽 [bit] / Bits per word
    DL_SHIFT32    : UDINT := 32;                       // 高字取回的固定移位量 [bit] / Fixed shift for the high word
END_VAR

(*------------------------------------------------------------------------------
 * 段 1｜输出预置：异常路径下全部输出确定
 *      Pre-set outputs so that every path is deterministic
 *-----------------------------------------------------------------------------*)
FC_DL_BitArrayInsert := FALSE;
nChanged             := 0;
uApplied             := 16#0000_0000_0000_0000;
uMask                := 16#0000_0000_0000_0000;
nActualW             := 0;
uErrorId             := 16#0000_0000;
bValid               := FALSE;

(*------------------------------------------------------------------------------
 * 段 2｜字数钳位与总位数（边界 B1）：先夹到 1 到 8
 *      Clamp the word count, then derive the total bit count
 *-----------------------------------------------------------------------------*)
IF nTargetCount < 1 THEN
    nTargetCount := 1;
ELSIF nTargetCount > DL_SRC_MAX THEN
    nTargetCount := DL_SRC_MAX;
END_IF
nTotalBits := INT_TO_DINT(nTargetCount) * INT_TO_DINT(DL_BIT_MAX32);

(*------------------------------------------------------------------------------
 * 段 3｜偏移闸门（边界 B2）：负偏移与落空偏移早退，绝不写半个字
 *      Offset gate: negative or beyond the stream end exits without writing
 *-----------------------------------------------------------------------------*)
IF (nOffset < 0) OR (INT_TO_DINT(nOffset) >= nTotalBits) THEN
    uErrorId := 16#0001_0128;   // 偏移越界，目标数组一字未动
    RETURN;
END_IF

(*------------------------------------------------------------------------------
 * 段 4｜宽度闸门（边界 B3）：宽度须落在 1 到 64 闭区间
 *      Width gate: the window width must be within one to sixty four
 *-----------------------------------------------------------------------------*)
IF (nWidth < 1) OR (nWidth > DL_BIT_MAX64) THEN
    uErrorId := 16#0001_0129;   // 宽度越界，目标数组一字未动
    RETURN;
END_IF

(*------------------------------------------------------------------------------
 * 段 5｜越界截断（边界 B4）：按位流末端截断，之后仍写可用低位
 *      Truncation at the stream end, the usable low bits are still written
 *-----------------------------------------------------------------------------*)
IF (INT_TO_DINT(nOffset) + INT_TO_DINT(nWidth)) > nTotalBits THEN
    nWidth   := DINT_TO_INT(nTotalBits - INT_TO_DINT(nOffset));
    uErrorId := 16#0001_012A;
    bValid   := FALSE;
END_IF

(*------------------------------------------------------------------------------
 * 段 6｜定位（边界 B5）：低字下标、字内移位量与跨字判据
 *      Locate the low word, the intra word shift and the straddle flag
 *-----------------------------------------------------------------------------*)
nIdxLo := nOffset / DL_BIT_MAX32 + 1;
nShift := nOffset MOD DL_BIT_MAX32;
nIdxHi := 0;
IF ((nShift + nWidth) > DL_BIT_MAX32) AND (nIdxLo < nTargetCount) THEN
    nIdxHi := nIdxLo + 1;
END_IF

(*------------------------------------------------------------------------------
 * 段 7｜双字窗口深度校验（边界 B6）：跨到第三个字时按双字窗口截断
 *      Third word guard: a window reaching the next word is truncated here
 *      起点非零时 64 位移位中间量只能覆盖到第二个字末尾，超出部分若继续写
 *      会把高位静默写成零，故显式截断并报事件
 *-----------------------------------------------------------------------------*)
IF (nShift + nWidth) > DL_BIT_MAX64 THEN
    nWidth   := DL_BIT_MAX64 - nShift;
    uErrorId := 16#0001_012A;
    bValid   := FALSE;
END_IF

(*------------------------------------------------------------------------------
 * 段 8｜掩码与生效值（边界 B7）：64 宽走常量分支，禁止左移 64 位
 *      Mask and applied value: the full width case uses the constant branch
 *-----------------------------------------------------------------------------*)
IF nWidth >= DL_BIT_MAX64 THEN
    uMask := DL_MASK64_ALL;
ELSE
    uMask := SHL(LWORD#1, INT_TO_UDINT(nWidth)) - LWORD#1;
END_IF
uApplied := uValue AND uMask;

(*------------------------------------------------------------------------------
 * 段 9｜展开到窗口位置：字内移位量 0 到 31，左移后必然落在 64 位内
 *      Shift mask and value up into the window position
 *      断言口径：段 6 与段 7 已保证移位量加宽度不超过 64，故此处不会溢出位宽
 *-----------------------------------------------------------------------------*)
uMaskWide := SHL(uMask, INT_TO_UDINT(nShift));
uWinWide  := SHL(uApplied, INT_TO_UDINT(nShift));

(*------------------------------------------------------------------------------
 * 段 10｜取旧值并逐字算出新值，此段只读不写
 *      Read the old words and compute the new ones, still no write here
 *-----------------------------------------------------------------------------*)
uOldLo := auTarget[nIdxLo];
uOldHi := 16#0000_0000;
IF nIdxHi > 0 THEN
    uOldHi := auTarget[nIdxHi];
END_IF
uNewLo := (uOldLo AND NOT LWORD_TO_DWORD(uMaskWide)) OR LWORD_TO_DWORD(uWinWide);
uNewHi := 16#0000_0000;
IF nIdxHi > 0 THEN
    uNewHi := (uOldHi AND NOT LWORD_TO_DWORD(SHR(uMaskWide, DL_SHIFT32))) OR LWORD_TO_DWORD(SHR(uWinWide, DL_SHIFT32));
END_IF

(*------------------------------------------------------------------------------
 * 段 11｜先比较后计数（边界 B8）：值未变的字不算改动，也不产生写动作
 *      Compare before counting: unchanged words are neither counted nor written
 *-----------------------------------------------------------------------------*)
IF uNewLo <> uOldLo THEN
    nChanged := nChanged + 1;
END_IF
IF (nIdxHi > 0) AND (uNewHi <> uOldHi) THEN
    nChanged := nChanged + 1;
END_IF

(*------------------------------------------------------------------------------
 * 段 12｜原子写回：新值全部算完之后再按低字、高字顺序落盘
 *      Atomic write back after all new values are known
 *      若值未变则跳过写动作，避免下游映像刷新产生无谓的总线负载
 *-----------------------------------------------------------------------------*)
IF uNewLo <> uOldLo THEN
    auTarget[nIdxLo] := uNewLo;
END_IF
IF (nIdxHi > 0) AND (uNewHi <> uOldHi) THEN
    auTarget[nIdxHi] := uNewHi;
END_IF

(*------------------------------------------------------------------------------
 * 段 13｜收口：宽度定稿，无事件时置有效与返回真
 *      Close out: publish the effective width, legal calls return true
 *-----------------------------------------------------------------------------*)
nActualW := nWidth;
IF uErrorId = 16#0000_0000 THEN
    bValid               := TRUE;
    FC_DL_BitArrayInsert := TRUE;
END_IF
END_FUNCTION

(* ---- FC_DL_BitArraySegCopy.st ---- *)
// =====================================================================
// FC_DL_BitArraySegCopy.st
// 位段数组多段一次搬（源到目标多段批量复制, 逐段域校验 + 整段原子性）
// Multi-segment batch bit-array copy with per-segment domain validation
// 所属子库: DL_Base    版本: v1.0.0    兼容: CODESYS V3.5+ / TwinCAT 3 / 汇川 InoProShop
// 码位: 16#0001_048E ~ 16#0001_0491 (本件独占 4 槽, FC 纯函数分型, 勿复用)
// 溯源: IEC 61131-3 标准语义的道莅防御性实现
//       来源组标签: bit-field, array-copy, batch-transfer, lgf-bitlogic
// 修改记录: R30 初版 (ROUND_PLAN_R30 序 20)
// 语义声明: 一次调用搬 N 段; 逐段域校验（起位 + 长度不超过数组位容量）
//           先整体校验后统一搬移, 任一段非法则零段搬移并回放段号;
//           跨字窗口逐位读改写沿用 Extract/Insert 范式（移位量以取余 32
//           归一, 全程仅 32 位移位, 无 64 位移位）; 段表内重叠段不做去重,
//           后段覆盖前段; 与 FC_DL_BitArrayExtract/Insert 逐段对拍位守恒
// =====================================================================
FUNCTION FC_DL_BitArraySegCopy : BOOL   // 返回真 = 全部段搬移完成 / TRUE when all segments copied
VAR_IN_OUT
    aSrc   : ARRAY[*] OF DWORD;     // 源位数组（开数组, 实测边界）/ Source bit array
    aDst   : ARRAY[*] OF DWORD;     // 目标位数组（开数组, 实测边界）/ Destination bit array
END_VAR
VAR_INPUT
    aSrcBit   : ARRAY[*] OF UINT;   // 各段源起始位号 0 起 / Per-segment source start bit
    aDstBit   : ARRAY[*] OF UINT;   // 各段目标起始位号 0 起 / Per-segment destination start bit
    aLen      : ARRAY[*] OF USINT;  // 各段长度（位）1~255 / Per-segment length in bits
    uSegCount : USINT;              // 段数 / Segment count
END_VAR
VAR_OUTPUT
    uErrorId : UDINT;               // 错误码, 见码表 / Error code, see table
    uFailSeg : USINT;               // 非法段号回放 1~N, 0 = 无 / Failed segment replay, 0 = none
END_VAR
VAR
    uSrcCap  : DINT := 0;           // 源数组实测位容量 / Source capacity in bits
    uDstCap  : DINT := 0;           // 目标数组实测位容量 / Destination capacity in bits
    uTabCap1 : DINT := 0;           // 段表 1 实测容量 / Segment table 1 capacity
    uTabCap2 : DINT := 0;           // 段表 2 实测容量 / Segment table 2 capacity
    uTabCap3 : DINT := 0;           // 段表 3 实测容量 / Segment table 3 capacity
    uTabCap  : DINT := 0;           // 段表最小容量 / Minimum table capacity
    uSegUse  : DINT := 0;           // 实际处理段数（钳位后）/ Effective segment count
    iS       : DINT := 0;           // 段循环下标 / Segment loop index
    iJ       : DINT := 0;           // 位循环下标 / Bit loop index
    iSIdx    : DINT := 0;           // 段表元素下标 / Segment table element index
    uSrcPos  : DINT := 0;           // 当前源位号 / Current source bit position
    uDstPos  : DINT := 0;           // 当前目标位号 / Current destination bit position
    iW       : DINT := 0;           // 字下标 / Word index
    dwMask   : DWORD := DWORD#0;    // 位掩码 / Bit mask
    dwWord   : DWORD := DWORD#0;    // 目标字读改写临时量 / Destination word read-modify-write temp
    xBit     : BOOL := FALSE;       // 当前位值 / Current bit value
    uSegLen  : DINT := 0;           // 当前段长度 / Current segment length
END_VAR

// ---------------------------------------------------------------------
// 代码位表（本件独占, 勿复用）:
//   16#0001_048E 信息 批量搬移完成（含段表重叠时后段覆盖前段语义）
//   16#0001_048F 信息 空段表（段数为 0, 零搬移成功返回）
//   16#0001_0490 故障 段域非法（起位 + 长度超过数组位容量, 段号经 uFailSeg
//                回放, 零段搬移原子回退）; 纯函数无锁存面, 修正段表重新调用即解除
//   16#0001_0491 信息 段计数越界钳位（段数大于段表实测容量, 已按容量截断处理）
// ---------------------------------------------------------------------

// ---- 缺省收口 / Defaults ----
FC_DL_BitArraySegCopy := FALSE;     // 缺省失败 / Default fail
uErrorId := 16#0001_048E;           // 缺省完成码, 异常路径覆盖 / Default done code
uFailSeg := 0;                      // 段号清零 / Clear segment number

// ---- 容量实测（开数组边界实测, 不假设下标起点）/ Measured capacities ----
uSrcCap := 32 * ((UPPER_BOUND(aSrc, 1) - LOWER_BOUND(aSrc, 1)) + 1);    // 源位容量 / Source bits
uDstCap := 32 * ((UPPER_BOUND(aDst, 1) - LOWER_BOUND(aDst, 1)) + 1);    // 目标位容量 / Destination bits
uTabCap1 := (UPPER_BOUND(aSrcBit, 1) - LOWER_BOUND(aSrcBit, 1)) + 1;
uTabCap2 := (UPPER_BOUND(aDstBit, 1) - LOWER_BOUND(aDstBit, 1)) + 1;
uTabCap3 := (UPPER_BOUND(aLen, 1) - LOWER_BOUND(aLen, 1)) + 1;
// 取三段表最小容量 / Minimum of the three table capacities
uTabCap := uTabCap1;
IF uTabCap2 < uTabCap THEN
    uTabCap := uTabCap2;
END_IF
IF uTabCap3 < uTabCap THEN
    uTabCap := uTabCap3;
END_IF

// ---- 空段表: 零搬移成功返回 / Empty segment table ----
IF uSegCount = 0 THEN
    uErrorId := 16#0001_048F;       // 空段表码 / Empty table code
    FC_DL_BitArraySegCopy := TRUE;  // 零搬移成功 / Zero-copy success
    RETURN;
END_IF

// ---- 段计数钳位（信息级, 按段表容量截断）/ Segment count clamp ----
uSegUse := USINT_TO_DINT(uSegCount);
IF uSegUse > uTabCap THEN
    uSegUse := uTabCap;             // 截断处理 / Truncate
    uErrorId := 16#0001_0491;       // 钳位信息码 / Clamp info code
END_IF

// ---- 整体校验: 逐段域校验, 任一非法即零段搬移退出（整段原子性）
//      Whole validation first, any invalid segment aborts with zero moved ----
FOR iS := 1 TO uSegUse DO
    iSIdx := LOWER_BOUND(aSrcBit, 1) + (iS - 1);    // 段表下标映射 / Table index mapping
    uSrcPos := UINT_TO_DINT(aSrcBit[iSIdx]);
    uSegLen := USINT_TO_DINT(aLen[iSIdx]);
    IF (uSrcPos + uSegLen) > uSrcCap THEN
        uErrorId := 16#0001_0490;   // 段域非法码 / Illegal segment domain
        uFailSeg := DINT_TO_USINT(iS);  // 回放段号 / Replay segment number
        RETURN;                     // 零段搬移退出 / Abort with zero moved
    END_IF
    uDstPos := UINT_TO_DINT(aDstBit[iSIdx]);
    IF (uDstPos + uSegLen) > uDstCap THEN
        uErrorId := 16#0001_0490;   // 段域非法码 / Illegal segment domain
        uFailSeg := DINT_TO_USINT(iS);
        RETURN;                     // 零段搬移退出 / Abort
    END_IF
END_FOR

// ---- 统一搬移: 逐段逐位读改写（后段覆盖前段, 不去重）/ Unified copy ----
FOR iS := 1 TO uSegUse DO
    iSIdx := LOWER_BOUND(aSrcBit, 1) + (iS - 1);
    uSegLen := USINT_TO_DINT(aLen[iSIdx]);
    uSrcPos := UINT_TO_DINT(aSrcBit[iSIdx]);    // 源位号复位 / Reset source position
    uDstPos := UINT_TO_DINT(aDstBit[iSIdx]);    // 目标位号复位 / Reset destination position
    FOR iJ := 1 TO uSegLen DO
        // 读源位（跨字窗口, 移位量取余 32 归一, 小于 32 位宽合规）
        // Read source bit across word boundary, shift normalized mod 32
        iW := LOWER_BOUND(aSrc, 1) + (uSrcPos / 32);
        dwMask := SHL(DWORD#1, uSrcPos MOD 32);
        xBit := (aSrc[iW] AND dwMask) <> DWORD#0;
        // 写目标位（读改写保持其余位）/ Write destination bit with read-modify-write
        iW := LOWER_BOUND(aDst, 1) + (uDstPos / 32);
        dwWord := aDst[iW];
        dwMask := SHL(DWORD#1, uDstPos MOD 32);
        IF xBit THEN
            dwWord := dwWord OR dwMask;             // 置位 / Set bit
        ELSE
            dwWord := dwWord AND (NOT dwMask);      // 清位 / Clear bit
        END_IF
        aDst[iW] := dwWord;                         // 回写字 / Write back
        uSrcPos := uSrcPos + 1;                     // 源位推进 / Advance source
        uDstPos := uDstPos + 1;                     // 目标位推进 / Advance destination
    END_FOR
END_FOR

FC_DL_BitArraySegCopy := TRUE;      // 全部段完成 / All segments done

END_FUNCTION

(* ---- FC_DL_BitCount.st ---- *)
(*==============================================================================
 * 组件名称 (Component)  : FC_DL_BitCount
 * 所属子库 (Sublibrary) : DL_Base
 * 当前版本 (Version)    : 1.0.0
 * 兼容性   (Platform)   : CODESYS 3.5 / TwinCAT 3 / 汇川 InoProShop / Machine Expert
 *                         仅用标准 AND / 减法 / WHILE，无任何厂商内建函数
 * 功能描述 (Function)   : 统计 32 位字中置 1 的位数（Hamming Weight / Population Count），
 *                         返回 0..32。用于多传感器投票表决、工位占用统计、报警字
 *                         严重度分级。采用 Brian Kernighan 法 uTemp AND (uTemp - 1)，
 *                         迭代次数等于置位数：全 0 输入零次、全 1 输入恰好 32 次，
 *                         避免逐位 FOR 的固定 32 次开销与差一错误。
 * 开源溯源 (Origin)     : 原创实现。Brian W. Kernighan 位计数法（公开经典算法，
 *                         见《The C Programming Language》习题 2-9），本处为 ST 重写。
 * 依赖     (Depends)    : 无 DL_ 内部依赖；无标准库功能块依赖
 * 红线自检 (Redline)    : R1 ✓ 零全局变量表与外部变量引用 ｜ R2 ✓ 零物理 IO 地址直写
 *                         R3 ✓ 纯 IEC 61131-3 ｜ R4 ✓ WHILE 防死锁计数器 + 无符号回绕前提注释
 *                         R5 ✓ 全变量中英双语同行注释 ｜ R6 N/A（无状态机）｜ R7 N/A（无实例调用）
 * 修订历史 (Revision)   :
 *   2026-11-14  v1.0.0  首版入库（Phase 1 冷启动 · Level 0 批次）
 *============================================================================*)
FUNCTION FC_DL_BitCount : USINT
VAR_INPUT
    uValue   : DWORD;    // 待统计的 32 位字 / 32-bit word to be counted
END_VAR
VAR_OUTPUT
    bValid   : BOOL;     // 计算完整标志，FALSE 表示触发循环保护 / Calculation complete flag, FALSE means loop guard tripped
    uErrorId : UDINT;    // 故障码，0 = 无故障 / Error code, 0 = no error
END_VAR
VAR
    uTemp    : DWORD;    // 工作副本，循环中被逐位清零 / Working copy, bits cleared one by one inside the loop
    nCount   : USINT;    // 置位计数，值域 0..32 / Population count, range 0..32
    nGuard   : DINT;     // 循环防死锁计数器 / Loop deadlock guard counter
END_VAR
VAR CONSTANT
    DL_POPCOUNT_MAX_LOOP : DINT := 32;  // 迭代上限，等于 Brian Kernighan 法的理论上界 / Iteration limit equal to the theoretical bound
END_VAR

(*------------------------------------------------------------------------------
 * 段 1｜返回值与工作变量初始化：任何路径下返回值确定
 *      Initialize return value and working variables for deterministic results
 *-----------------------------------------------------------------------------*)
FC_DL_BitCount := 16#00;
bValid         := TRUE;
uErrorId       := 16#0000_0000;
uTemp          := uValue;
nCount         := 16#00;
nGuard         := 0;

(*------------------------------------------------------------------------------
 * 段 2｜Brian Kernighan 位计数（边界 B1/B2/B3）
 *      Brian Kernighan population count (boundaries B1/B2/B3)
 *      每次 uTemp AND (uTemp - 1) 精确清除最低位的 1，迭代次数 = 置位数
 *      前提：uTemp - 1 的无符号回绕仅在 uTemp 非零时安全，故"非零"写进
 *            WHILE 条件成为循环不变式，而非仅写在注释里的口头约定
 *      Premise: the unsigned wrap of (uTemp - 1) is safe only while uTemp <> 0,
 *               therefore the non-zero test lives in the WHILE condition itself
 *-----------------------------------------------------------------------------*)
WHILE (uTemp <> 16#0000_0000) AND (nGuard < DL_POPCOUNT_MAX_LOOP) DO
    uTemp  := uTemp AND (uTemp - 16#0000_0001);
    nCount := nCount + 16#01;
    nGuard := nGuard + 1;
END_WHILE;

(*------------------------------------------------------------------------------
 * 段 3｜循环完整性判定（边界 B2）
 *      Loop completeness check (boundary B2)
 *      判据取"残值是否归零"而非"计数器是否到顶"：全 1 输入在第 32 次迭代
 *      同时使残值归零与计数器到顶，若只比对计数器会误报循环保护
 *      The residual value is the criterion, not the guard counter: an all-ones
 *      input reaches both limits simultaneously and would be falsely flagged
 *-----------------------------------------------------------------------------*)
IF uTemp <> 16#0000_0000 THEN
    bValid   := FALSE;
    uErrorId := 16#0001_0004;
END_IF

(*------------------------------------------------------------------------------
 * 段 4｜结果回写（边界 B4/B5）：USINT 容量 255 远大于 32，无溢出风险
 *      Result write-back: USINT capacity 255 far exceeds 32, overflow impossible
 *-----------------------------------------------------------------------------*)
FC_DL_BitCount := nCount;
END_FUNCTION

(* ---- FC_DL_BitCountOnes.st ---- *)
(*
  Name        : FC_DL_BitCountOnes
  Category    : DL_Base
  Version     : 1.0.0
  Purpose     : 位串置 1 计数（popcount）：逐位单热掩码扫描统计 DWORD 中为 1 的位数，输出 0..32；/ Population count of set bits in a DWORD, walking-one mask scan, result 0..32
  溯源        : 借 t2-1-lgf·bitlogic 的分类/参数域组织，clean-room 实现
  Boundary    : ① 位宽固定 32 位（DWORD 为跨平台最宽公共无符号型；LWORD 64 位需平台确认，本族另件）；
                ② 移位量恒 0..31 < 32，绝不出现 SHL(x, 位宽) 的未定义行为（末拍 SHL(16#80000000,1)=0 无害）；
                ③ 输出域钳位 0..32，防越界写入下游；
                ④ 输入 NaN 概念不适用（整型），无除零路径（纯位运算）。
*)
FUNCTION FC_DL_BitCountOnes : INT
VAR_INPUT
    dwBits     : DWORD := 0;                 (* 待计数位串，按 32 位解释 [-] / Bit string to count, 32-bit *)
    xEarlyExit : BOOL := TRUE;               (* 提前退出：剩余未扫描位已全 0 时终止循环（省周期）[-] / Early exit when remaining bits are zero *)
END_VAR
VAR
    dwMask : DWORD;                          (* 逐位单热掩码，初值 1 后每拍左移 1 位 [-] / Walking-one mask *)
    dwRest : DWORD;                          (* 剩余未扫描位串（早退出判据）[-] / Remaining unscanned bits *)
    nIdx   : INT;                            (* 位序号游标 0..31（FOR 自复位，R227）[-] / Bit index cursor 0..31 *)
    nAcc   : INT;                            (* 累加计数 0..32 [-] / Accumulated count 0..32 *)
END_VAR
VAR CONSTANT
    DL_BCO_WIDTH : INT   := 32;              (* DWORD 位宽（移位量上界基准，恒 < 本值）[位] / DWORD bit width *)
    DL_BCO_MAX   : INT   := 32;              (* 计数结果上限（防越界，R308）[位] / Count result ceiling *)
    DL_BCO_ONE   : DWORD := 1;               (* 单热掩码初值（最低位置 1）[-] / Initial walking-one mask *)
    DL_BCO_ZERO  : DWORD := 0;               (* 位串零常量（比较用，避免魔法数）[-] / Zero constant for comparison *)
END_VAR

(* —— 段 1：单拍量预清零（R107：每拍全路径派生，无跨拍残留） —— *)
nAcc := 0;                                   (* 累加器预清 / Accumulator preset *)
dwMask := DL_BCO_ONE;                        (* 掩码回到最低位 / Mask to LSB *)
dwRest := dwBits;                            (* 剩余位串取输入全量 / Remaining bits = input *)

(* —— 段 2：逐位扫描（FOR 上限 < 位宽，移位量归一，R28） —— *)
FOR nIdx := 0 TO DL_BCO_WIDTH - 1 DO
    IF (dwRest = DL_BCO_ZERO) AND xEarlyExit THEN
        EXIT;                                (* 剩余位全 0：提前终止，计数已定 / Early exit, count settled *)
    END_IF
    IF (dwBits AND dwMask) <> DL_BCO_ZERO THEN
        nAcc := nAcc + 1;                     (* 该位为 1：计数递增 / Bit set: increment *)
    END_IF
    dwRest := dwRest AND NOT dwMask;          (* 清除已扫描位（NOT 为按位取反，DWORD 语义） / Clear scanned bit *)
    dwMask := SHL(dwMask, 1);                 (* 掩码左移一位（1..31 < 32，无越界） / Shift mask left, amount < width *)
END_FOR

(* —— 段 3：输出饱和（硬限反算：极限值 32 为 INT 可表，安全） —— *)
IF nAcc < 0 THEN
    nAcc := 0;                                (* 下限兜底（理论不可达，防御性） / Lower bound fallback *)
ELSIF nAcc > DL_BCO_MAX THEN
    nAcc := DL_BCO_MAX;                       (* 上限饱和 32 [位] / Upper saturation to 32 *)
END_IF
FC_DL_BitCountOnes := nAcc;                  (* 函数返回：置 1 位数 / Return: number of set bits *)
END_FUNCTION
